(* IEC 61131-3 sources: PLC-IsaVODE/PLC-IsaVODE/samples/plc-programs (part 13) *)

(* ---- 727-SNTP_CLIENT.ST ---- *)
TYPE
  oscat_IP_FIFO128_DATA  : ARRAY [1..128] OF BYTE;
  oscat_Mailbox  : ARRAY [1..16] OF BYTE;

  oscat_IP_FIFO_DATA :
  STRUCT
    X       : oscat_IP_FIFO128_DATA; (* IP_ID FIFO Speicher          *)
    Y       : oscat_IP_FIFO128_DATA; (* IP_ID Z�hler                 *)
    ID      : BYTE;                  (* h�chste vergabene id         *)
    MAX_ID  : BYTE;                  (* maximal Anmeldungen pro ID   *)
      INIT    : BOOL;                  (* Initialisierung durchgef�hrt *)
    EMPTY   : BOOL;                  (* FIFO leer                    *)
    FULL    : BOOL;                  (* FIFO voll                    *)
    TOP     : INT;                   (* maximale anzahl in FIFO      *)
    NW      : INT;                   (* Schreibzeiger                *)
    NR      : INT;                   (* Lesezeiger                   *)
  END_STRUCT;

  oscat_IP_C:
  STRUCT
    C_MODE:			BYTE;          		(*W Mode: TCP/UCP AKTIV/PASSIV                               *)
    C_PORT:         WORD;          		(*W Portnummer                                               *)
    C_IP:           DWORD;         		(*W IP-Adresse gepackt wwxxyyzz = www.xxx.yyy.zzz            *)
    C_STATE:        BYTE;          		(*R Verbindungsstatus ON/OFF + Flanke ON/OFF                 *)
    C_ENABLE:       BOOL;          		(*W Freigabe f�r Connect                                     *)
    R_OBSERVE:      BOOL;          		(*W Empfang ueberwachen                                      *)
    TIME_RESET:     BOOL;          		(*W Alle Timer ruecksetzen                                   *)
    ERROR:          DWORD;         		(*R vvwwxxyy (vv = CON_ERROR, ww = SEN_ERROR, xx = REC_ERROR *)
    FIFO:           oscat_IP_FIFO_DATA; (*I IP FIFO Struktur                                         *)
    MAILBOX:		oscat_Mailbox;		(*I Mailbox: Datenbereich f�r Bausteindatenaustausch         *)
  END_STRUCT;
END_TYPE

TYPE

  oscat_NW_BUF_LONG  : ARRAY [0..4095] OF BYTE;

  oscat_NETWORK_BUFFER :
  STRUCT
    SIZE   : UINT;
    BUFFER : oscat_NW_BUF_LONG;
  END_STRUCT;

END_TYPE

FUNCTION _BYTE_TO_INT:INT
	VAR_INPUT
		IN :	BYTE;
	END_VAR

	_BYTE_TO_INT := USINT_TO_INT(BYTE_TO_USINT(IN));
END_FUNCTION

FUNCTION_BLOCK IP_FIFO_Block

  VAR_IN_OUT
    FIFO :	oscat_IP_FIFO_DATA;
    ID :	BYTE;
    STATE :	BYTE;
  END_VAR

  VAR
    tmp :	INT;
  END_VAR

  IF NOT FIFO.INIT THEN
    FIFO.INIT		:= TRUE;
    FIFO.NW		:= 1;
    FIFO.NR		:= 1;
    FIFO.EMPTY	:= TRUE;
    FIFO.FULL		:= FALSE;
    FIFO.TOP		:= 128;
    FIFO.MAX_ID	:= BYTE#1;
  END_IF;

  IF ID = BYTE#00 THEN
    IF FIFO.ID < INT_TO_BYTE(FIFO.TOP) THEN
      ID := USINT_TO_BYTE(BYTE_TO_USINT(FIFO.ID) + USINT#1);
      FIFO.ID := ID ;

    ELSIF STATE < BYTE#200 THEN
      STATE := BYTE#255;
    RETURN;
    END_IF;
  END_IF;

  IF STATE = BYTE#1 AND NOT FIFO.FULL THEN
    tmp := _BYTE_TO_INT(ID);
    IF FIFO.Y[tmp] < FIFO.MAX_ID THEN
      FIFO.Y[tmp] := USINT_TO_BYTE(BYTE_TO_USINT(FIFO.Y[tmp]) + USINT#1);
      tmp := FIFO.NW;
      FIFO.X[tmp] := ID;
      IF FIFO.NW = FIFO.TOP THEN FIFO.NW := 1; ELSE FIFO.NW := FIFO.NW + 1; END_IF;
      FIFO.FULL := FIFO.NW = FIFO.NR;
    FIFO.EMPTY := FALSE;
      STATE := BYTE#2;
    END_IF;
  END_IF;

  IF STATE = BYTE#2 AND NOT FIFO.EMPTY THEN
    tmp := FIFO.NR;
    IF ID = FIFO.X[tmp] THEN
      STATE := BYTE#3;
    END_IF;
  END_IF;

  IF STATE = BYTE#4 AND NOT FIFO.EMPTY THEN

    tmp := FIFO.NR;
    IF ID = FIFO.X[tmp] THEN
      tmp := _BYTE_TO_INT(ID);
      FIFO.Y[tmp] := USINT_TO_BYTE(BYTE_TO_USINT(FIFO.Y[tmp]) - USINT#1);

      IF FIFO.NR = FIFO.TOP THEN FIFO.NR := 1; ELSE FIFO.NR := FIFO.NR + 1; END_IF;
      FIFO.EMPTY := FIFO.NR = FIFO.NW;
    FIFO.FULL := FALSE;
    END_IF;
    STATE := BYTE#5;
  END_IF;

END_FUNCTION_BLOCK

FUNCTION_BLOCK T_PLC_MS_block

	VAR_OUTPUT
		T_PLC_MS :	UDINT;
	END_VAR

	VAR_EXTERNAL
		PLC_TICKS_PER_SEC :	INT;
		PLC_SYS_TICK_CNT :	DINT;
	END_VAR

	VAR
		debug :	BOOL;(*Debug-Mode ON / OFF*)
		N :	INT;(*Debug-Faktor*)
		Offset :	UDINT;(*Debug-Offset*)
		temp :	DWORD := DWORD#1;(*Debug-Offset*)
		mode :	BOOL;(*modus*)
		faktor :	UDINT;(*Systemtakt-Faktor*)
		init :	BOOL;
		v_plc_ticks_per_sec :	UDINT;
		base :	UDINT := UDINT#1000;
	END_VAR

	IF init = FALSE THEN
		v_plc_ticks_per_sec := INT_TO_UDINT(PLC_TICKS_PER_SEC);
		IF v_plc_ticks_per_sec = UDINT#1024 THEN
			faktor := UDINT#1;
			mode := FALSE;
		ELSIF v_plc_ticks_per_sec > UDINT#0 THEN
			IF v_plc_ticks_per_sec <= base THEN
				faktor := base / v_plc_ticks_per_sec;
				mode := FALSE;
			ELSE
				faktor := v_plc_ticks_per_sec / base;
				mode := TRUE;
			END_IF;
		ELSE
			faktor := UDINT#1;
		END_IF;
		init := TRUE;
	END_IF;

	IF mode THEN
		T_PLC_MS := DINT_TO_UDINT(PLC_SYS_TICK_CNT) / faktor;
	ELSE
		T_PLC_MS := DINT_TO_UDINT(PLC_SYS_TICK_CNT) * faktor;
	END_IF;

	IF debug THEN
		T_PLC_MS := (DWORD_TO_UDINT(SHL(UDINT_TO_DWORD(T_PLC_MS),N) OR SHL(temp,N)) - UDINT#1) + Offset;
	END_IF;

END_FUNCTION_BLOCK

FUNCTION DWORD_OF_BYTE:DWORD
	VAR_INPUT
		B3 :	BYTE;
		B2 :	BYTE;
		B1 :	BYTE;
		B0 :	BYTE;
	END_VAR

	DWORD_OF_BYTE := SHL(SHL(SHL(BYTE_TO_DWORD(B3),8) OR BYTE_TO_DWORD(B2),8) OR BYTE_TO_DWORD(B1),8) OR BYTE_TO_DWORD(B0);

END_FUNCTION

FUNCTION _WORD_TO_DINT:DINT
	VAR_INPUT
		IN :	WORD;
	END_VAR
	_WORD_TO_DINT := UINT_TO_DINT(WORD_TO_UINT(IN));
END_FUNCTION

FUNCTION WORD_OF_BYTE:WORD
	VAR_INPUT
		B1 :	BYTE;
		B0 :	BYTE;
	END_VAR
	WORD_OF_BYTE := SHL(BYTE_TO_WORD(B1),8) OR BYTE_TO_WORD(B0);
END_FUNCTION

FUNCTION _INT_TO_UDINT:UDINT
	VAR_INPUT
		IN :	INT;
	END_VAR

	_INT_TO_UDINT := DINT_TO_UDINT(INT_TO_DINT(IN));
END_FUNCTION

FUNCTION_BLOCK SNTP_CLIENT_Block

  VAR_IN_OUT
    IP_C :	oscat_IP_C;
    S_BUF :	oscat_NETWORK_BUFFER;
    R_BUF :	oscat_NETWORK_BUFFER;
  END_VAR

  VAR_INPUT
    IP4 :	DWORD;
    ACTIVATE :	BOOL;
  END_VAR

  VAR_OUTPUT
    ERROR :	DWORD;
    DONE_P :	BOOL;
    UDT :	UDINT;
    XMS :	INT;
  END_VAR

  VAR
    IP_STATE :	BYTE;
    IP_ID :	BYTE;
    IP_FIFO :	IP_FIFO_Block;
    i :	INT;
    last :	UDINT;
    state :	INT;
    T_PLC_MS :	T_PLC_MS_Block;
    tx :	UDINT;
    ACTIVATE_LAST :	BOOL;
    IP4_STORED :	DWORD;
  END_VAR

  T_PLC_MS();
  tx := T_PLC_MS.T_PLC_MS;

  CASE state OF
  00:
    DONE_P := FALSE;
    IF ACTIVATE AND NOT ACTIVATE_LAST THEN
      IP4_STORED := IP4;
      state := 10;
      ERROR := DWORD#0;
      IP_STATE := BYTE#1;
    END_IF;

  10:
    IF IP_STATE = BYTE#3 THEN

      S_BUF.BUFFER[00] := BYTE#16#1B;
      FOR i := 1 TO 47 DO
        S_BUF.BUFFER[i] := BYTE#16#00;
      END_FOR;

      last := tx;
      state := 30;

      IP_C.C_PORT     := WORD#123;
      IP_C.C_IP       := IP4_STORED;
      IP_C.C_MODE     := BYTE#1;
      IP_C.C_ENABLE   := TRUE;
      IP_C.TIME_RESET := TRUE;
      IP_C.R_OBSERVE  := TRUE;
      S_BUF.SIZE      := UINT#48;
      R_BUF.SIZE      := UINT#0;
    END_IF;

  30:
    IF IP_C.ERROR <> DWORD#00 THEN
      ERROR := IP_C.ERROR;
    S_BUF.SIZE := UINT#0;
    R_BUF.SIZE := UINT#0;
      state := 0;
    ELSIF S_BUF.SIZE = UINT#0 AND R_BUF.SIZE >= UINT#48 THEN
      UDT := DWORD_TO_UDINT(DWORD_OF_BYTE(R_BUF.BUFFER[40],R_BUF.BUFFER[41],R_BUF.BUFFER[42],R_BUF.BUFFER[43]))- UDINT#2208988800;

      XMS := DWORD_TO_INT(SHR(DINT_TO_DWORD(_WORD_TO_DINT(WORD_OF_BYTE(R_BUF.BUFFER[44],R_BUF.BUFFER[45])) * DINT#1000),16));
      XMS := XMS + DWORD_TO_INT(SHR(UDINT_TO_DWORD(tx - last),1));

      UDT := UDT + _INT_TO_UDINT(XMS / 1000);
      XMS := XMS MOD 1000;

      state := 0;
      DONE_P := TRUE;

    END_IF;

    IF state = 0 THEN
      IP_C.R_OBSERVE := FALSE;
      IP_STATE := BYTE#4;
    END_IF;

  END_CASE;

  ACTIVATE_LAST := ACTIVATE;

  IP_FIFO(FIFO:=IP_C.FIFO,STATE:=IP_STATE,ID:=IP_ID);
  IP_C.FIFO:=IP_FIFO.FIFO;
  IP_STATE := IP_FIFO.STATE;
  IP_ID:=IP_FIFO.ID;

END_FUNCTION_BLOCK

PROGRAM program0
	VAR
		IP_C :	oscat_IP_C;
    S_BUF :	oscat_NETWORK_BUFFER;
    R_BUF :	oscat_NETWORK_BUFFER;
    IP4 :	DWORD;
    ACTIVATE :	BOOL;
    ERROR :	DWORD;
    DONE_P :	BOOL;
    UDT :	UDINT;
    XMS :	INT;

		func_block : SNTP_CLIENT_Block;
	END_VAR
	func_block.IP_C := IP_C;
	func_block.S_BUF := S_BUF;
	func_block.R_BUF := R_BUF;
  func_block.IP4 := IP4;
	func_block.ACTIVATE := ACTIVATE;

	func_block();
  IP_C  := func_block.IP_C;
  S_BUF  := func_block.S_BUF;
  R_BUF  := func_block.R_BUF;
  ERROR  := func_block.ERROR;
  DONE_P  := func_block.DONE_P;
  UDT  := func_block.UDT;
  XMS  := func_block.XMS;
END_PROGRAM

CONFIGURATION Config0

	VAR_GLOBAL
		PLC_TICKS_PER_SEC :	INT;
		PLC_SYS_TICK_CNT :	DINT;
	END_VAR

  	RESOURCE Res0 ON PLC
    	TASK task0(INTERVAL := T#20ms,PRIORITY := 0);
    	PROGRAM instance0 WITH task0 : program0;
  	END_RESOURCE

END_CONFIGURATION

(* ---- 728-HOLIDAY.ST ---- *)
TYPE oscat_LANGUAGE:
  STRUCT
    DEFAULT 	: INT;
	LMAX    	: INT;
  END_STRUCT;
END_TYPE

TYPE
	oscat_LOCATION_ELEMENTS	: ARRAY [1..5] OF INT;
END_TYPE

TYPE
  oscat_ELEMENT_WEEKDAYS	: ARRAY [1..7] OF STRING;
  oscat_WEEKDAYS			: ARRAY [1..3]  OF oscat_ELEMENT_WEEKDAYS := [0, 0, 0];
END_TYPE

TYPE oscat_LOCATION:
  STRUCT
    DEFAULT 	: INT;
	LMAX    	: INT;
	LANGUAGE	: oscat_LOCATION_ELEMENTS;
  END_STRUCT;
END_TYPE

TYPE oscat_HOLIDAY_DATA :
  STRUCT
	NAME : STRING;
	DAY : SINT;
	MONTH : SINT;
	USE : SINT;
	PAD_BYTE : BYTE;
  END_STRUCT;
END_TYPE

TYPE
  oscat_HOLIDAY_DATA_0_29 	: ARRAY [0..29] OF oscat_HOLIDAY_DATA;
  oscat_HOLIDAY_DATA_0_49 	: ARRAY [0..49] OF oscat_HOLIDAY_DATA;
END_TYPE

FUNCTION_BLOCK SETUP_LANGUAGE_Block

	VAR_IN_OUT
		LANGUAGE :	oscat_LANGUAGE;
	END_VAR

	VAR
		init :	BOOL;
	END_VAR

	IF init THEN RETURN; END_IF;
	init := TRUE;

	LANGUAGE.DEFAULT  := 1; (* 1=english, 2=german 3=french *)
	LANGUAGE.LMAX := 3;
END_FUNCTION_BLOCK

FUNCTION_BLOCK SETUP_LOCATION
	VAR_IN_OUT
		LOCATION :	oscat_LOCATION;
	END_VAR

	VAR
		init :	BOOL;
	END_VAR

	IF init THEN RETURN; END_IF;
	init := TRUE;

	LOCATION.DEFAULT  := 1;
	LOCATION.LMAX := 5;

	LOCATION.LANGUAGE[1] := 2;
	LOCATION.LANGUAGE[2] := 2;
	LOCATION.LANGUAGE[3] := 3;
	LOCATION.LANGUAGE[4] := 2;
	LOCATION.LANGUAGE[5] := 2;
END_FUNCTION_BLOCK

FUNCTION_BLOCK SETUP_WEEKDAYS

	VAR_IN_OUT
		WEEKDAYS :	oscat_WEEKDAYS;
	END_VAR

	VAR
		init :	BOOL;
	END_VAR

	IF init THEN RETURN; END_IF;
	init := TRUE;

	WEEKDAYS[1][01] := 'Monday';
	WEEKDAYS[1][02] := 'Tuesday';
	WEEKDAYS[1][03] := 'Wednesday';
	WEEKDAYS[1][04] := 'Thursday';
	WEEKDAYS[1][05] := 'Friday';
	WEEKDAYS[1][06] := 'Saturday';
	WEEKDAYS[1][07] := 'Sunday';

	WEEKDAYS[2][01] := 'Montag';
	WEEKDAYS[2][02] := 'Dienstag';
	WEEKDAYS[2][03] := 'Mittwoch';
	WEEKDAYS[2][04] := 'Donnerstag';
	WEEKDAYS[2][05] := 'Freitag';
	WEEKDAYS[2][06] := 'Samstag';
	WEEKDAYS[2][07] := 'Sonntag';

	WEEKDAYS[3][01] := 'Lundi';
	WEEKDAYS[3][02] := 'Mardi';
	WEEKDAYS[3][03] := 'Mercredi';
	WEEKDAYS[3][04] := 'Jeudi';
	WEEKDAYS[3][05] := 'Vendredi';
	WEEKDAYS[3][06] := 'Samedi';
	WEEKDAYS[3][07] := 'Dimanche';
END_FUNCTION_BLOCK

FUNCTION YEAR_OF_DATE:INT
	VAR_INPUT
		IDATE :	UDINT;
	END_VAR

	YEAR_OF_DATE := UDINT_TO_INT((idate+UDINT#43200) / UDINT#31557600 + UDINT#1970);
END_FUNCTION

FUNCTION _INT_TO_UDINT:UDINT
	VAR_INPUT
		IN :	INT;
	END_VAR

	_INT_TO_UDINT := DINT_TO_UDINT(INT_TO_DINT(IN));
END_FUNCTION

FUNCTION SET_DATE:UDINT

	VAR_INPUT
		YEAR :	INT;
		MONTH :	INT;
		DAY :	INT;
	END_VAR

	VAR
		count :	INT;
	END_VAR

	IF month > 2 THEN
		count := (month - 1) * 30;
		IF month > 7 THEN
			count := count + DWORD_TO_INT(SHR(DINT_TO_DWORD(INT_TO_DINT(month) - INT_TO_DINT(3)),1));
		ELSE
			count := count + DWORD_TO_INT(SHR(DINT_TO_DWORD(INT_TO_DINT(month) - INT_TO_DINT(4)),1));
		END_IF;
		IF SHL(INT_TO_WORD(year),14) = WORD#0 THEN
			count := count + 1;
		END_IF;
	ELSE
		count := (month - 1) * 31;
	END_IF;
	SET_DATE := (_INT_TO_UDINT(count + day - 1) + DWORD_TO_UDINT(SHR(UDINT_TO_DWORD(_INT_TO_UDINT(year) * UDINT#1461 - UDINT#2878169), 2))) * UDINT#86400;
END_FUNCTION

FUNCTION DAY_OF_WEEK:INT
	VAR_INPUT
		IDATE :	UDINT;
	END_VAR

	DAY_OF_WEEK := UDINT_TO_INT((idate / UDINT#86400 + UDINT#3) MOD UDINT#7) + INT#01;
END_FUNCTION

FUNCTION EASTER:UDINT
	VAR_INPUT
		YEAR :	INT;
	END_VAR

	VAR
		b :	INT;
		c :	INT;
		oday :	INT;
	END_VAR

	b := (204 - 11 * (year MOD 19)) MOD 30;
	IF b > 27 THEN b := b - 1; END_IF;
	c := (year + WORD_TO_INT(SHR(INT_TO_WORD(year),2)) + b - 13) MOD 7;
	oday := 28 + b - c;
	IF oday > 33 THEN
		easter := set_Date(year, 4, oday - 31);
	ELSE
		easter := set_Date(year, 3, oday);
	END_IF;
END_FUNCTION

FUNCTION LEAP_OF_DATE:BOOL

	VAR_INPUT
		IDATE :	UDINT;
	END_VAR

	LEAP_OF_DATE := SHL(UDINT_TO_DWORD((idate + UDINT#43200) / UDINT#31557600), 30) = DWORD#16#80000000;
END_FUNCTION

FUNCTION DAY_OF_YEAR:INT
	VAR_INPUT
		IDATE :	UDINT;
	END_VAR

	DAY_OF_YEAR := UDINT_TO_INT(((idate) / UDINT#86400) MOD UDINT#1461);
	IF DAY_OF_YEAR > 729 THEN
		IF DAY_OF_YEAR > 1095 THEN DAY_OF_YEAR := DAY_OF_YEAR - 1095; ELSE DAY_OF_YEAR := DAY_OF_YEAR - 729; END_IF;
	ELSIF DAY_OF_YEAR > 364 THEN
		DAY_OF_YEAR := DAY_OF_YEAR - 364;
	ELSE
		DAY_OF_YEAR := DAY_OF_YEAR + 1;
	END_IF;
END_FUNCTION

FUNCTION MONTH_OF_DATE:INT

	VAR_INPUT
		IDATE :	UDINT;
	END_VAR

	MONTH_OF_DATE := DAY_OF_YEAR(idate);
	IF MONTH_OF_DATE < 32 THEN
		MONTH_OF_DATE := 1;
	ELSIF LEAP_OF_DATE((IDATE)) THEN
		MONTH_OF_DATE := (MONTH_OF_DATE * 53 + 1668) / 1623;
	ELSE
		MONTH_OF_DATE := (MONTH_OF_DATE * 53 + 1700) / 1620;
	END_IF;
END_FUNCTION

FUNCTION DAY_OF_MONTH:INT
	VAR_INPUT
		IDATE :	UDINT;
	END_VAR

	day_of_month := day_of_year(idate);

	IF leap_of_Date((idate)) THEN
		CASE day_of_month OF
			32..60	:	day_of_month := day_of_month - 31;
			61..91	:	day_of_month := day_of_month - 60;
			92..121 :	day_of_month := day_of_month - 91;
			122..152:	day_of_month := day_of_month - 121;
			153..182:	day_of_month := day_of_month - 152;
			183..213:	day_of_month := day_of_month - 182;
			214..244:	day_of_month := day_of_month - 213;
			245..274:	day_of_month := day_of_month - 244;
			275..305:	day_of_month := day_of_month - 274;
			306..335:	day_of_month := day_of_month - 305;
			336..366:	day_of_month := day_of_month - 335;
		END_CASE;
	ELSE
		CASE day_of_month OF
			32..59	:	day_of_month := day_of_month - 31;
			60..90	:	day_of_month := day_of_month - 59;
			91..120 :	day_of_month := day_of_month - 90;
			121..151:	day_of_month := day_of_month - 120;
			152..181:	day_of_month := day_of_month - 151;
			182..212:	day_of_month := day_of_month - 181;
			213..243:	day_of_month := day_of_month - 212;
			244..273:	day_of_month := day_of_month - 243;
			274..304:	day_of_month := day_of_month - 273;
			305..334:	day_of_month := day_of_month - 304;
			335..365:	day_of_month := day_of_month - 334;
		END_CASE;
	END_IF;
END_FUNCTION

FUNCTION DATE_ADD:UDINT
	VAR_INPUT
		IDATE :	UDINT;
		D :	INT;
		W :	INT;
		M :	INT;
		Y :	INT;
	END_VAR

	VAR
		mo :	INT;
		yr :	INT;
		dm :	INT;
	END_VAR

	DATE_ADD := IDATE + INT_TO_UDINT(D + W * 7) * UDINT#86400;
	yr := Y + YEAR_OF_DATE(DATE_ADD);
	mo := M + MONTH_OF_DATE(DATE_ADD);
	dm := DAY_OF_MONTH(DATE_ADD);
	WHILE mo > 12 DO
		mo := mo - 12;
		yr := yr + 1;
	END_WHILE;
	WHILE mo < 1 DO
		mo := mo + 12;
		yr := yr - 1;
	END_WHILE;
	DATE_ADD := SET_DATE(yr, mo, dm);
END_FUNCTION

FUNCTION_BLOCK HOLIDAY_Block
	VAR_INPUT
		DATE_IN :	UDINT;
		LANGU :	INT;
		FRIDAY :	BOOL;
		SATURDAY :	BOOL;
		SUNDAY :	BOOL;
	END_VAR

	VAR_IN_OUT
		HOLIDAYS :	oscat_HOLIDAY_DATA_0_29;
	END_VAR

	VAR_OUTPUT
		Y :	BOOL;
		NAME :	STRING;
	END_VAR

	VAR
		size :	INT := INT#29;
		last_active :	UDINT;
		ostern :	UDINT;
		i :	INT;
		jahr :	INT;
		x_date :	UDINT;
		lx :	INT;
		wdx :	INT;
		SETUP_LOCATIONS :	SETUP_LOCATION;
		SETUP_WEEKDAYSS :	SETUP_WEEKDAYS;
		SETUP_LANGUAGES :	SETUP_LANGUAGE_Block;
		LOCATION :	oscat_LOCATION;
		WEEKDAYS :	oscat_WEEKDAYS;
		LANGUAGE :	oscat_LANGUAGE;
		wd :	INT;
	END_VAR

	IF last_active = date_in THEN RETURN; END_IF;
	last_active := DATE_IN;

	SETUP_LOCATIONS(LOCATION:=LOCATION);
	LOCATION:=SETUP_LOCATIONS.LOCATION;

	SETUP_WEEKDAYSS(WEEKDAYS:=WEEKDAYS);
	WEEKDAYS:=SETUP_WEEKDAYSS.WEEKDAYS;

	SETUP_LANGUAGES(LANGUAGE:=LANGUAGE);
	LANGUAGE:=SETUP_LANGUAGES.LANGUAGE;

	IF LANGU = 0 THEN
		lx := language.DEFAULT;
	ELSE
		lx := MIN(language.LMAX, LANGU);
	END_IF;

	jahr := YEAR_OF_DATE(date_in);
	ostern := EASTER(jahr);
	wdx := DAY_OF_WEEK(DATE_IN);
	Y := FALSE;

	FOR i := 0 TO size DO
		x_date := SET_DATE(jahr, SINT_TO_INT(HOLIDAYS[i].MONTH) , SINT_TO_INT(HOLIDAYS[i].DAY));
		IF HOLIDAYS[i].USE = SINT#1 AND HOLIDAYS[i].MONTH > SINT#0 THEN
			(* check for fixed date holiday *)
			IF x_date = date_in THEN
				Y := TRUE;
				NAME := HOLIDAYS[i].NAME;
				RETURN;
			END_IF;
		ELSIF HOLIDAYS[i].USE = SINT#1 AND HOLIDAYS[i].MONTH = SINT#0 THEN
			(* check for holiday in reference to easter *)
			IF DATE_ADD(ostern, SINT_TO_INT(HOLIDAYS[i].DAY),0,0,0) = date_in THEN
				Y := TRUE;
				NAME := HOLIDAYS[i].NAME;
				RETURN;
			END_IF;
		ELSIF HOLIDAYS[i].USE < SINT#0 THEN
			(* check for holiday on a weekday before date *)
			IF DAY_OF_WEEK(date_in) = SINT_TO_INT(ABS(HOLIDAYS[i].USE)) AND date_in < x_date AND date_in >= DATE_ADD(x_date,-7,0,0,0) THEN
				Y := TRUE;
				NAME := HOLIDAYS[i].NAME;
				RETURN;
			END_IF;
		END_IF;
	END_FOR;

	IF NOT Y AND (wdx = 5 AND FRIDAY OR wdx = 6 AND SATURDAY OR wdx = 7 AND SUNDAY) THEN
		Y := TRUE;
		wd := LOCATION.LANGUAGE[lx];
		NAME := WEEKDAYS[wd][wdx];
	ELSE
		NAME := '';
	END_IF;
END_FUNCTION_BLOCK

PROGRAM program0
  VAR
	DATE_IN  :	UDINT;
	LANGU    :	INT;
	FRIDAY   :	BOOL;
	SATURDAY :	BOOL;
	SUNDAY   :	BOOL;

	Y :	BOOL;
	NAME :	STRING;

	HOLIDAYS :	oscat_HOLIDAY_DATA_0_29;

	func_block : HOLIDAY_Block;
  END_VAR
	func_block.DATE_IN :=DATE_IN ;
	func_block.LANGU   :=LANGU   ;
	func_block.FRIDAY  :=FRIDAY  ;
	func_block.SATURDAY:=SATURDAY;
	func_block.SUNDAY  :=SUNDAY  ;
	func_block.HOLIDAYS  :=HOLIDAYS ;

	func_block();
	Y := func_block.Y;
	NAME := func_block.NAME;
	HOLIDAYS := func_block.HOLIDAYS;

END_PROGRAM

CONFIGURATION Config0
  RESOURCE Res0 ON PLC
    TASK task0(INTERVAL := T#20ms,PRIORITY := 0);
    PROGRAM instance0 WITH task0 : program0;
  END_RESOURCE
END_CONFIGURATION

(* ---- 732-LEGIONELLA.ST ---- *)
FUNCTION TIMECHECK:BOOL

	VAR_INPUT
		TD :	UDINT;
		START :	UDINT;
		STOP :	UDINT;
	END_VAR

	IF stop < start THEN
		TIMECHECK := start <= TD OR  TD < stop;
	ELSE
		TIMECHECK := start <= TD AND TD < stop;
	END_IF;

END_FUNCTION

FUNCTION TIME_TO_TOD:UDINT

	VAR_INPUT
		IN :	TIME;
	END_VAR

	TIME_TO_TOD := DWORD_TO_UDINT(TIME_TO_DWORD(IN));
END_FUNCTION

FUNCTION TOD_TO_TIME:TIME
	VAR_INPUT
		IN :	UDINT;
	END_VAR

	TOD_TO_TIME := DWORD_TO_TIME(UDINT_TO_DWORD(IN));
END_FUNCTION

FUNCTION DAY_OF_WEEK:INT
  VAR_INPUT
    IDATE :	UDINT;
  END_VAR

  DAY_OF_WEEK := UDINT_TO_INT((idate / UDINT#86400 + UDINT#3) MOD UDINT#7) + INT#01;
END_FUNCTION

FUNCTION _DT_TO_DATE_B:UDINT

	VAR_INPUT
		_INN :	UDINT;
	END_VAR

	_DT_TO_DATE_B := (_INN / UDINT#86400) * UDINT#86400;
END_FUNCTION

FUNCTION DT_TO_TOD2:UDINT
	VAR_INPUT
		IN :	UDINT;
	END_VAR

	DT_TO_TOD2 := (IN MOD UDINT#86400) * UDINT#1000;
END_FUNCTION

FUNCTION TIME_TO_TOD2:UDINT

	VAR_INPUT
		IN :	TIME;
	END_VAR

	TIME_TO_TOD2 := DWORD_TO_UDINT(TIME_TO_DWORD(IN));
END_FUNCTION

FUNCTION_BLOCK TIMER_1_Block

	VAR_INPUT
		E :	BOOL := TRUE;
		DTI :	UDINT;
		START :	UDINT;
		DURATION :	TIME;
		DAY :	BYTE := BYTE#2#0111_1111;
	END_VAR

	VAR_OUTPUT
		Q :	BOOL;
		STOP :	TIME;
	END_VAR

	IF E THEN
		stop := TOD_TO_TIME(START) + DURATION;
		IF stop > T#24h THEN stop := stop - T#24h; END_IF;
		Q := TIMECHECK(DT_TO_TOD2(DTI), START, TIME_TO_TOD2(stop)) AND (SHR(BYTE#128, DAY_OF_WEEK(_DT_TO_DATE_B(DTI))) AND DAY) > BYTE#0;
	ELSE
		Q := FALSE;
	END_IF;

END_FUNCTION_BLOCK

FUNCTION UDINT_TO_TIME2:TIME

	VAR_INPUT
		IN :	UDINT;
	END_VAR

	UDINT_TO_TIME2 := DINT_TO_TIME(UDINT_TO_DINT(IN));

END_FUNCTION

FUNCTION_BLOCK T_PLC_MS_block
	VAR_OUTPUT
		T_PLC_MS :	UDINT;
	END_VAR

	VAR_EXTERNAL
		PLC_TICKS_PER_SEC :	INT;
		PLC_SYS_TICK_CNT :	DINT;
	END_VAR

	VAR
		debug :	BOOL;
		N :	INT;
		Offset :	UDINT;
		temp :	DWORD := DWORD#1;
		mode :	BOOL;
		faktor :	UDINT;
		init :	BOOL;
		v_plc_ticks_per_sec :	UDINT;
		base :	UDINT := UDINT#1000;
	END_VAR

	IF init = FALSE THEN
		v_plc_ticks_per_sec := INT_TO_UDINT(PLC_TICKS_PER_SEC);
		IF v_plc_ticks_per_sec = UDINT#1024 THEN
			faktor := UDINT#1;
			mode := FALSE;
		ELSIF v_plc_ticks_per_sec > UDINT#0 THEN
			IF v_plc_ticks_per_sec <= base THEN
				faktor := base / v_plc_ticks_per_sec;
				mode := FALSE;
			ELSE
				faktor := v_plc_ticks_per_sec / base;
				mode := TRUE;
			END_IF;
		ELSE
			faktor := UDINT#1;
		END_IF;
		init := TRUE;
	END_IF;

	IF mode THEN
		T_PLC_MS := DINT_TO_UDINT(PLC_SYS_TICK_CNT) / faktor;
	ELSE
		T_PLC_MS := DINT_TO_UDINT(PLC_SYS_TICK_CNT) * faktor;
	END_IF;

	IF debug THEN
		T_PLC_MS := (DWORD_TO_UDINT(SHL(UDINT_TO_DWORD(T_PLC_MS),N) OR SHL(temp,N)) - UDINT#1) + Offset;
	END_IF;

END_FUNCTION_BLOCK

FUNCTION_BLOCK SEQUENCE_8_Block

	VAR_INPUT
		IN0 :	BOOL := TRUE;
		IN1 :	BOOL := TRUE;
		IN2 :	BOOL := TRUE;
		IN3 :	BOOL := TRUE;
		IN4 :	BOOL := TRUE;
		IN5 :	BOOL := TRUE;
		IN6 :	BOOL := TRUE;
		IN7 :	BOOL := TRUE;
		START :	BOOL;
		RST :	BOOL;
		WAIT0 :	TIME;
		DELAY0 :	TIME;
		WAIT1 :	TIME;
		DELAY1 :	TIME;
		WAIT2 :	TIME;
		DELAY2 :	TIME;
		WAIT3 :	TIME;
		DELAY3 :	TIME;
		WAIT4 :	TIME;
		DELAY4 :	TIME;
		WAIT5 :	TIME;
		DELAY5 :	TIME;
		WAIT6 :	TIME;
		DELAY6 :	TIME;
		WAIT7 :	TIME;
		DELAY7 :	TIME;
		STOP_ON_ERROR :	BOOL;
	END_VAR

	VAR_OUTPUT
		Q0 :	BOOL;
		Q1 :	BOOL;
		Q2 :	BOOL;
		Q3 :	BOOL;
		Q4 :	BOOL;
		Q5 :	BOOL;
		Q6 :	BOOL;
		Q7 :	BOOL;
		QX :	BOOL;
		RUN :	BOOL;
		_STEP :	INT := -1;
		STATUS :	BYTE;
	END_VAR

	VAR
		last :	TIME;
		edge :	BOOL;
		tx :	TIME;
		init :	BOOL;
		T_PLC_MS :	T_PLC_MS_Block;
	END_VAR

	T_PLC_MS();
	tx:= UDINT_TO_TIME(T_PLC_MS.T_PLC_MS);

	IF NOT init THEN
		last := tx;
		init := TRUE;
		status := BYTE#110;
	END_IF;

	IF rst THEN
		_step := -1;
		Q0 := FALSE;
		Q1 := FALSE;
		Q2 := FALSE;
		Q3 := FALSE;
		Q4 := FALSE;
		Q5 := FALSE;
		Q6 := FALSE;
		Q7 := FALSE;
		status := BYTE#110;
		run := FALSE;

	ELSIF start AND NOT edge THEN
		_step := 0;
		last := tx;
		status := BYTE#111;
		Q0 := FALSE;
		Q1 := FALSE;
		Q2 := FALSE;
		Q3 := FALSE;
		Q4 := FALSE;
		Q5 := FALSE;
		Q6 := FALSE;
		Q7 := FALSE;
		run := TRUE;
	END_IF;
	edge := start;

	IF status > BYTE#0 AND status < BYTE#100 AND stop_on_error THEN RETURN; END_IF;

	IF run AND _step = 0 THEN
		IF NOT q0 AND in0 AND tx - last <= wait0 THEN
			Q0 := TRUE;
			last := tx;
		ELSIF NOT q0 AND tx - last > wait0 THEN
			status := BYTE#1;
			run := FALSE;
		ELSIF q0 AND tx - last >= delay0 THEN
			_step := 1;
			last := tx;
		END_IF;
	END_IF;
	IF run AND _step = 1 THEN
		IF NOT q1 AND in1 AND tx - last <= wait1 THEN
			Q0 := FALSE;
			Q1 := TRUE;
			last := tx;
		ELSIF NOT q1 AND Tx - last > wait1 THEN
			status := BYTE#2;
			q0 := FALSE;
			run := FALSE;
		ELSIF q1 AND tx - last >= delay1 THEN
			_step := 2;
			last := tx;
		END_IF;
	END_IF;
	IF run AND _step = 2 THEN
		IF NOT q2 AND in2 AND tx - last <= wait2 THEN
			Q1 := FALSE;
			Q2 := TRUE;
			last := tx;
		ELSIF NOT q2 AND Tx - last > wait2 THEN
			status := BYTE#3;
			q1 := FALSE;
			run := FALSE;
		ELSIF q2 AND tx - last >= delay2 THEN
			_step := 3;
			last := tx;
		END_IF;
	END_IF;
	IF run AND _step = 3 THEN
		IF NOT q3 AND in3 AND tx - last <= wait3 THEN
			Q2 := FALSE;
			Q3 := TRUE;
			last := tx;
		ELSIF NOT q3 AND Tx - last > wait3 THEN
			status := BYTE#4;
			q2 := FALSE;
			run := FALSE;
		ELSIF q3 AND tx - last >= delay3 THEN
			_step := 4;
			last := tx;
		END_IF;
	END_IF;
	IF run AND _step = 4 THEN
		IF NOT q4 AND in4 AND tx - last <= wait4 THEN
			Q3 := FALSE;
			Q4 := TRUE;
			last := tx;
		ELSIF NOT q4 AND Tx - last > wait4 THEN
			status := BYTE#5;
			q3 := FALSE;
			run := FALSE;
		ELSIF q4 AND tx - last >= delay4 THEN
			_step := 5;
			last := tx;
		END_IF;
	END_IF;
	IF run AND _step = 5 THEN
		IF NOT q5 AND in5 AND tx - last <= wait5 THEN
			Q4 := FALSE;
			Q5 := TRUE;
			last := tx;
		ELSIF NOT q5 AND Tx - last > wait5 THEN
			status := BYTE#6;
			q4 := FALSE;
			run := FALSE;
		ELSIF q5 AND tx - last >= delay5 THEN
			_step := 6;
			last := tx;
		END_IF;
	END_IF;
	IF run AND _step = 6 THEN
		IF NOT q6 AND in6 AND tx - last <= wait6 THEN
			Q5 := FALSE;
			Q6 := TRUE;
			last := tx;
		ELSIF NOT q6 AND Tx - last > wait6 THEN
			status := BYTE#7;
			q5 := FALSE;
			run := FALSE;
		ELSIF q6 AND tx - last >= delay6 THEN
			_step := 7;
			last := tx;
		END_IF;
	END_IF;
	IF run AND _step = 7 THEN
		IF NOT q7 AND in7 AND tx - last <= wait7 THEN
			Q6 := FALSE;
			Q7 := TRUE;
			last := tx;
		ELSIF NOT q7 AND Tx - last > wait7 THEN
			status := BYTE#8;
			q6 := FALSE;
			run := FALSE;
		ELSIF q7 AND tx - last >= delay7 THEN
			_step := -1;
			Q7 := FALSE;
			Run := FALSE;
			status := BYTE#110;
		END_IF;
	END_IF;
	QX := q0 OR q1 OR q2 OR q3 OR q4 OR q5 OR q6 OR q7;

END_FUNCTION_BLOCK

FUNCTION_BLOCK HYST_1_Block

	VAR_INPUT
		IN :	REAL;
		HIGH :	REAL;
		LOW :	REAL;
	END_VAR

	VAR_OUTPUT
		Q :	BOOL;
		WIN :	BOOL;
	END_VAR

	IF in < low THEN
		Q := FALSE;
		win := FALSE;
	ELSIF in > high THEN
		Q := TRUE;
		win := FALSE;
	ELSE
		win := TRUE;
	END_IF;

END_FUNCTION_BLOCK

FUNCTION_BLOCK LEGIONELLA_Block

	VAR_INPUT
		MANUAL :	BOOL;
		TEMP_BOILER :	REAL;
		TEMP_RETURN :	REAL := 100.0;
		DT_IN :	UDINT;
		RST :	BOOL;
		T_START :	UDINT := UDINT#10800000;(*tod#03:00:00*)
		DAY :	INT := 7;
		TEMP_SET :	REAL := 70.0;
		TEMP_OFFSET :	REAL := 10.0;
		TEMP_HYS :	REAL := 5.0;
		T_MAX_HEAT :	TIME := t#10m;
		T_MAX_RET :	TIME := t#10m;
		TP_0 :	TIME := t#5m;
		TP_1 :	TIME := t#5m;
		TP_2 :	TIME := t#5m;
		TP_3 :	TIME := t#5m;
		TP_4 :	TIME := t#5m;
		TP_5 :	TIME := t#5m;
		TP_6 :	TIME := t#5m;
		TP_7 :	TIME := t#5m;
	END_VAR

	VAR_OUTPUT
		HEAT :	BOOL;
		PUMP :	BOOL;
		VALVE0 :	BOOL;
		VALVE1 :	BOOL;
		VALVE2 :	BOOL;
		VALVE3 :	BOOL;
		VALVE4 :	BOOL;
		VALVE5 :	BOOL;
		VALVE6 :	BOOL;
		VALVE7 :	BOOL;
		RUN :	BOOL;
		_STATUS :	BYTE;
	END_VAR

	VAR
		X1 :	TIMER_1_Block;
		x2 :	SEQUENCE_8_Block;
		x3 :	HYST_1_Block;
		init :	BOOL;
	END_VAR

	IF NOT init THEN
		init := TRUE;
		X1.day := SHR(BYTE#128,day);
		X1.start := T_start;
		X3.low := Temp_offset + temp_set;
		X3.high := Temp_hys + X3.low;
		X2.wait0 := T_max_heat;
		X2.delay0 := TP_0;
		X2.delay1 := TP_1;
		X2.delay2 := TP_2;
		X2.delay3 := TP_3;
		X2.delay4 := TP_4;
		X2.delay5 := TP_5;
		X2.delay6 := TP_6;
		X2.delay7 := TP_7;
		X2.wait1 := T_max_ret;
		X2.wait2 := T_max_ret;
		X2.wait3 := T_max_ret;
		X2.wait4 := T_max_ret;
		X2.wait5 := T_max_ret;
		X2.wait6 := T_max_ret;
		X2.wait7 := T_max_ret;
		X2();
	END_IF;

	X1(DTi := DT_in);
	IF X1.Q OR MANUAL OR x2.run THEN
		X3(in := temp_boiler);
		X2.in0 := X3.Q OR x3.win;
		X2.in1 := temp_return >= temp_set;
		X2.in2 := x2.in1;
		X2.in3 := x2.in1;
		X2.in4 := x2.in1;
		X2.in5 := x2.in1;
		X2.in6 := x2.in1;
		X2.in7 := x2.in1;
		X2.rst := rst;
		X2(start := X1.Q OR MANUAL);
		run := x2.run;
		pump := x2.QX;
		Heat := NOT X3.Q AND x2.run;
		valve0 := X2.Q0;
		valve1 := X2.Q1;
		valve2 := X2.Q2;
		valve3 := X2.Q3;
		valve4 := X2.Q4;
		valve5 := X2.Q5;
		valve6 := X2.Q6;
		valve7 := X2.Q7;
		pump := X2.QX;
		_STATUS := X2.status;
	ELSE
		X2(start := FALSE);
		_STATUS := x2.status;
	END_IF;

END_FUNCTION_BLOCK

PROGRAM program0
	VAR
		MANUAL :	BOOL;
		TEMP_BOILER :	REAL;
		TEMP_RETURN :	REAL := 100.0;
		DT_IN :	UDINT;
		RST :	BOOL;
		T_START :	UDINT := UDINT#10800000;(*tod#03:00:00*)
		DAY :	INT := 7;
		TEMP_SET :	REAL := 70.0;
		TEMP_OFFSET :	REAL := 10.0;
		TEMP_HYS :	REAL := 5.0;
		T_MAX_HEAT :	TIME := t#10m;
		T_MAX_RET :	TIME := t#10m;
		TP_0 :	TIME := t#5m;
		TP_1 :	TIME := t#5m;
		TP_2 :	TIME := t#5m;
		TP_3 :	TIME := t#5m;
		TP_4 :	TIME := t#5m;
		TP_5 :	TIME := t#5m;
		TP_6 :	TIME := t#5m;
		TP_7 :	TIME := t#5m;
		HEAT :	BOOL;
		PUMP :	BOOL;
		VALVE0 :	BOOL;
		VALVE1 :	BOOL;
		VALVE2 :	BOOL;
		VALVE3 :	BOOL;
		VALVE4 :	BOOL;
		VALVE5 :	BOOL;
		VALVE6 :	BOOL;
		VALVE7 :	BOOL;
		RUN :	BOOL;
		_STATUS :	BYTE;

		func_block : LEGIONELLA_Block;
	END_VAR
	func_block.MANUAL := MANUAL;
	func_block.TEMP_BOILER := TEMP_BOILER;
	func_block.TEMP_RETURN := TEMP_RETURN ;
	func_block.DT_IN    := DT_IN    ;
	func_block.RST := RST;
	func_block.T_START := T_START;
	func_block.DAY := DAY ;
	func_block.TEMP_SET := TEMP_SET ;
	func_block.TEMP_OFFSET    := TEMP_OFFSET    ;
	func_block.TEMP_HYS    := TEMP_HYS    ;
	func_block.T_MAX_HEAT := T_MAX_HEAT;
	func_block.T_MAX_RET := T_MAX_RET;
	func_block.TP_0 := TP_0;
	func_block.TP_1 := TP_1 ;
	func_block.TP_2 := TP_2 ;
	func_block.TP_3    := TP_3    ;
	func_block.TP_4    := TP_4    ;
	func_block.TP_5 := TP_5;
	func_block.TP_6 := TP_6;
	func_block.TP_7 := TP_7;

	func_block();
	HEAT  := func_block.HEAT;
	PUMP  := func_block.PUMP;
	VALVE0  := func_block.VALVE0;
	VALVE1  := func_block.VALVE1;
	VALVE2  := func_block.VALVE2;
	VALVE3  := func_block.HEAT;
	VALVE4  := func_block.VALVE4;
	VALVE5  := func_block.VALVE5;
	VALVE6  := func_block.VALVE6;
	VALVE7  := func_block.VALVE7;
	RUN  := func_block.RUN;
	_status  := func_block._status;
END_PROGRAM

CONFIGURATION Config0
	VAR_GLOBAL
		PLC_TICKS_PER_SEC :	INT;
		PLC_SYS_TICK_CNT :	DINT;
	END_VAR
  	RESOURCE Res0 ON PLC
    	TASK task0(INTERVAL := T#20ms,PRIORITY := 0);
    	PROGRAM instance0 WITH task0 : program0;
  	END_RESOURCE
END_CONFIGURATION

(* ---- 734-DCF77.ST ---- *)
TYPE
  oscat_dcf77_bits            : ARRAY [0..58]   OF BOOL;
END_TYPE

FUNCTION_BLOCK T_PLC_MS_block
	VAR_OUTPUT
		T_PLC_MS :	UDINT;
	END_VAR

	VAR_EXTERNAL
		PLC_TICKS_PER_SEC :	INT;
		PLC_SYS_TICK_CNT :	DINT;
	END_VAR

	VAR
		debug :	BOOL;(*Debug-Mode ON / OFF*)
		N :	INT;(*Debug-Faktor*)
		Offset :	UDINT;(*Debug-Offset*)
		temp :	DWORD := DWORD#1;(*Debug-Offset*)
		mode :	BOOL;(*modus*)
		faktor :	UDINT;(*Systemtakt-Faktor*)
		init :	BOOL;
		v_plc_ticks_per_sec :	UDINT;
		base :	UDINT := UDINT#1000;
	END_VAR

	IF init = FALSE THEN
		v_plc_ticks_per_sec := INT_TO_UDINT(PLC_TICKS_PER_SEC);
		IF v_plc_ticks_per_sec = UDINT#1024 THEN
			faktor := UDINT#1;
			mode := FALSE;
		ELSIF v_plc_ticks_per_sec > UDINT#0 THEN
			IF v_plc_ticks_per_sec <= base THEN
				faktor := base / v_plc_ticks_per_sec;
				mode := FALSE;
			ELSE
				faktor := v_plc_ticks_per_sec / base;
				mode := TRUE;
			END_IF;
		ELSE
			faktor := UDINT#1;
		END_IF;
		init := TRUE;
	END_IF;

	IF mode THEN
		T_PLC_MS := DINT_TO_UDINT(PLC_SYS_TICK_CNT) / faktor;
	ELSE
		T_PLC_MS := DINT_TO_UDINT(PLC_SYS_TICK_CNT) * faktor;
	END_IF;

	IF debug THEN
		T_PLC_MS := (DWORD_TO_UDINT(SHL(UDINT_TO_DWORD(T_PLC_MS),N) OR SHL(temp,N)) - UDINT#1) + Offset;
	END_IF;

END_FUNCTION_BLOCK

FUNCTION BIT_LOAD_W:WORD
	VAR_INPUT
		IN :	WORD;
		VAL :	BOOL;
		POS :	INT;
	END_VAR

	IF VAL THEN
		BIT_LOAD_W := in OR SHL(WORD#1,pos);
	ELSE
		BIT_LOAD_W := in AND (NOT SHL(WORD#1,pos));
	END_IF;
END_FUNCTION

FUNCTION BIT_OF_DWORD:BOOL
	VAR_INPUT
		IN :	DWORD;
		N :	INT;
	END_VAR
	BIT_OF_DWORD := (SHR(in,n) AND DWORD#1) > DWORD#0;
END_FUNCTION

FUNCTION EVEN:BOOL
	VAR_INPUT
		IN :	DINT;
	END_VAR
	even := NOT BIT_OF_DWORD(DINT_TO_DWORD(in),0);
END_FUNCTION

FUNCTION _INT_TO_UDINT:UDINT
	VAR_INPUT
		IN :	INT;
	END_VAR

	_INT_TO_UDINT := DINT_TO_UDINT(INT_TO_DINT(IN));
END_FUNCTION

FUNCTION SET_DATE:UDINT

	VAR_INPUT
		YEAR :	INT;
		MONTH :	INT;
		DAY :	INT;
	END_VAR

	VAR
		count :	INT;
	END_VAR

	IF month > 2 THEN
		count := (month - 1) * 30;
		IF month > 7 THEN
			count := count + DWORD_TO_INT(SHR(DINT_TO_DWORD(INT_TO_DINT(month) - INT_TO_DINT(3)),1));
		ELSE
			count := count + DWORD_TO_INT(SHR(DINT_TO_DWORD(INT_TO_DINT(month) - INT_TO_DINT(4)),1));
		END_IF;
		IF SHL(INT_TO_WORD(year),14) = WORD#0 THEN
			count := count + 1;
		END_IF;
	ELSE
		count := (month - 1) * 31;
	END_IF;
	SET_DATE := (_INT_TO_UDINT(count + day - 1) + DWORD_TO_UDINT(SHR(UDINT_TO_DWORD(_INT_TO_UDINT(year) * UDINT#1461 - UDINT#2878169), 2))) * UDINT#86400;

END_FUNCTION

FUNCTION DST:BOOL
	VAR_INPUT
		UTC :	UDINT;
	END_VAR

	VAR
		yr :	INT;
		yr4 :	UDINT;
		ltc :	UDINT;
		idate :	UDINT;
	END_VAR

	yr := YEAR_OF_DATE(DT_TO_DATE2(UTC));
	ltc := UTC;
	idate := SET_DT(yr, 3, 31, 1, 0, 0);
	yr4 := DWORD_TO_UDINT(SHR(INT_TO_DWORD(5 * yr), 2)) + UDINT#1;
	DST := (idate - ((yr4 + UDINT#3) MOD UDINT#7) * UDINT#86400 <= ltc) AND (idate + (UDINT#214 - (yr4) MOD UDINT#7) * UDINT#86400 > ltc);

END_FUNCTION

FUNCTION YEAR_OF_DATE:INT
	VAR_INPUT
		IDATE :	UDINT;
	END_VAR

	YEAR_OF_DATE := UDINT_TO_INT((idate+UDINT#43200) / UDINT#31557600 + UDINT#1970);
END_FUNCTION

FUNCTION DAY_OF_WEEK:INT

	VAR_INPUT
		IDATE :	UDINT;
	END_VAR

	DAY_OF_WEEK := UDINT_TO_INT((idate / UDINT#86400 + UDINT#3) MOD UDINT#7) + INT#01;
END_FUNCTION

FUNCTION SET_DT:UDINT
	VAR_INPUT
		YEAR :	INT;
		MONTH :	INT;
		DAY :	INT;
		HOUR :	INT;
		MINUTE :	INT;
		SECOND :	INT;
	END_VAR

	SET_DT := SET_DATE(YEAR, MONTH, DAY) + _INT_TO_UDINT(SECOND) + _INT_TO_UDINT(MINUTE) * UDINT#60 + _INT_TO_UDINT(HOUR) * UDINT#3600;
END_FUNCTION

FUNCTION DT_TO_DATE2:UDINT

	VAR_INPUT
		IN :	UDINT;
	END_VAR

	DT_TO_DATE2 := (IN / UDINT#86400) * UDINT#86400;

END_FUNCTION

FUNCTION_BLOCK DCF77
	VAR_INPUT
		REC :	BOOL;
		SET :	BOOL;
		SDT :	UDINT;
		DSI :	BOOL;
		SYNC_TIMEOUT :	TIME := t#2m;
		TIME_OFFSET :	INT := 1;
		DST_EN :	BOOL := TRUE;
	END_VAR

	VAR_OUTPUT
		TPp :	BOOL;
		DS :	BOOL;
		WDAY :	INT;
		ERROR :	BOOL;
		RTC2 :	UDINT;
		RTC21 :	UDINT;
		MSEC :	INT;
		SYNC :	BOOL;
	END_VAR

	VAR
		MEZ :	UDINT;
		UTC :	UDINT;
		state :	INT;
		edge :	BOOL;
		tx :	TIME;
		ty :	TIME;
		last :	TIME;
		bits :	oscat_dcf77_bits;
		cnt :	INT;
		i :	INT;
		old_time :	UDINT;
		minute :	INT;
		hour :	INT;
		day :	INT;
		month :	INT;
		year :	INT;
		last_sync :	TIME;
		t1 :	TIME;
		tz :	TIME;
		init :	BOOL;
		word_temp :	WORD;
		bool_temp :	BOOL;
		T_PLC_MS :	T_PLC_MS_block;
	END_VAR

	TPp := FALSE;

	T_PLC_MS();
	t1:= UDINT_TO_TIME(T_PLC_MS.T_PLC_MS);
	tx := t1 - last;

	IF rec XOR edge THEN
		edge := rec;
		IF NOT rec AND tx > t#1700ms AND tx < t#2000ms THEN
			(* start condition reached *)
			state := 0;
			tpp := NOT error;
		ELSIF NOT rec AND tx > t#700ms AND tx < t#1000ms THEN
			(* second switch detected *)
			IF state < 58 THEN state := state +1; ELSE state := 0; END_IF;
		ELSIF rec AND tx  < t#120ms THEN
			(* bit 0 detected  *)
			bits[state] := FALSE;
		ELSIF rec AND tx > t#120ms AND tx < t#250ms THEN
			(* bit 1 detected *)
			bits[state] := TRUE;
		ELSE
			(* error condition received signal is not valid *)
			error := TRUE;
			state := 0;
		END_IF;
		last := last + tx;
		IF rec AND state = 58 THEN
			error := FALSE;

			IF bits[0] OR NOT (bits[17] XOR bits[18]) OR NOT bits[20] THEN error := TRUE; END_IF;
			word_temp := WORD#0;

			bool_temp:=bits[21];
			word_temp:=BIT_LOAD_W(word_temp,bool_temp,0);
			bool_temp:=bits[22];
			word_temp:=BIT_LOAD_W(word_temp,bool_temp,1);
			bool_temp:=bits[23];
			word_temp:=BIT_LOAD_W(word_temp,bool_temp,2);
			bool_temp:=bits[24];
			word_temp:=BIT_LOAD_W(word_temp,bool_temp,3);

			minute := WORD_TO_INT(word_temp);
			IF bits[25] THEN minute := minute +10; END_IF;
			IF bits[26] THEN minute := minute +20; END_IF;
			IF bits[27] THEN minute := minute +40; END_IF;
			IF minute > 59 OR (bits[21] XOR bits[22] XOR bits[23] XOR bits[24] XOR bits[25] XOR bits[26] XOR bits[27] XOR bits[28]) THEN error := TRUE; END_IF;

			(* decode hour *)
			word_temp := WORD#0;

			bool_temp:=bits[29];
			word_temp:=BIT_LOAD_W(word_temp,bool_temp,0);    (* word_temp.X0 := bits[29]; *)
			bool_temp:=bits[30];
			word_temp:=BIT_LOAD_W(word_temp,bool_temp,1);    (* word_temp.X1 := bits[30]; *)
			bool_temp:=bits[31];
			word_temp:=BIT_LOAD_W(word_temp,bool_temp,2);    (* word_temp.X2 := bits[31]; *)
			bool_temp:=bits[32];
			word_temp:=BIT_LOAD_W(word_temp,bool_temp,3);    (* word_temp.X3 := bits[32]; *)

			hour := WORD_TO_INT(word_temp);
			IF bits[33] THEN hour := hour +10; END_IF;
			IF bits[34] THEN hour := hour +20; END_IF;
			IF hour > 23 OR (bits[29] XOR bits[30] XOR bits[31] XOR bits[32] XOR bits[33] XOR bits[34] XOR bits[35]) THEN error := TRUE; END_IF;

			(* decode day of month *)
			word_temp := WORD#0;

			bool_temp:=bits[36];
			word_temp:=BIT_LOAD_W(word_temp,bool_temp,0);    (* word_temp.X0 := bits[36]; *)
			bool_temp:=bits[37];
			word_temp:=BIT_LOAD_W(word_temp,bool_temp,1);    (* word_temp.X1 := bits[37]; *)
			bool_temp:=bits[38];
			word_temp:=BIT_LOAD_W(word_temp,bool_temp,2);    (* word_temp.X2 := bits[38]; *)
			bool_temp:=bits[39];
			word_temp:=BIT_LOAD_W(word_temp,bool_temp,3);    (* word_temp.X3 := bits[39]; *)

			day := WORD_TO_INT(word_temp);
			IF bits[40] THEN day := day + 10; END_IF;
			IF bits[41] THEN day := day + 20; END_IF;
			IF day > 31 THEN error := TRUE; END_IF;

			(* decode day of week *)
			word_temp := WORD#0;

			bool_temp:=bits[42];
			word_temp:=BIT_LOAD_W(word_temp,bool_temp,0);    (* word_temp.X0 := bits[42]; *)
			bool_temp:=bits[43];
			word_temp:=BIT_LOAD_W(word_temp,bool_temp,1);    (* word_temp.X1 := bits[43]; *)
			bool_temp:=bits[44];
			word_temp:=BIT_LOAD_W(word_temp,bool_temp,2);    (* word_temp.X2 := bits[44]; *)

			wday := WORD_TO_INT(word_temp);
			IF wday > 7 OR wday < 1 THEN error := TRUE; END_IF;

			(* decode month *)
			word_temp := WORD#0;

			bool_temp:=bits[45];
			word_temp:=BIT_LOAD_W(word_temp,bool_temp,0);    (* word_temp.X0 := bits[45]; *)
			bool_temp:=bits[46];
			word_temp:=BIT_LOAD_W(word_temp,bool_temp,1);    (* word_temp.X1 := bits[46]; *)
			bool_temp:=bits[47];
			word_temp:=BIT_LOAD_W(word_temp,bool_temp,2);    (* word_temp.X2 := bits[47]; *)
			bool_temp:=bits[48];
			word_temp:=BIT_LOAD_W(word_temp,bool_temp,3);    (* word_temp.X3 := bits[48]; *)

			month := WORD_TO_INT(word_temp);
			IF bits[49] THEN month := month +10; END_IF;
			IF month > 12 THEN error := TRUE; END_IF;

			(* decode year *)
			word_temp := WORD#0;

			bool_temp:=bits[50];
			word_temp:=BIT_LOAD_W(word_temp,bool_temp,0);    (* word_temp.X0 := bits[50]; *)
			bool_temp:=bits[51];
			word_temp:=BIT_LOAD_W(word_temp,bool_temp,1);    (* word_temp.X1 := bits[51]; *)
			bool_temp:=bits[52];
			word_temp:=BIT_LOAD_W(word_temp,bool_temp,2);    (* word_temp.X2 := bits[52]; *)
			bool_temp:=bits[53];
			word_temp:=BIT_LOAD_W(word_temp,bool_temp,3);    (* word_temp.X3 := bits[53]; *)

			year := WORD_TO_INT(word_temp);
			IF bits[54] THEN year := year + 10; END_IF;
			IF bits[55] THEN year := year + 20; END_IF;
			IF bits[56] THEN year := year + 40; END_IF;
			IF bits[57] THEN year := year + 80; END_IF;

			(* check parity for bits 36 to 58 *)
			cnt := 0;
			FOR i := 36 TO 58 DO IF bits[i] THEN cnt := cnt + 1; END_IF; END_FOR;
			IF NOT even(INT_TO_DINT(cnt)) THEN error := TRUE; END_IF;

			(* time must be valid for two cycles to clear error flag *)
			IF NOT error THEN
				(* set outputs *)
				old_time := mez;
				IF year >= 70 THEN year := year + 1900; ELSE year := year + 2000; END_IF;
				mez := set_DT(year,month,day,hour,minute,0);
				DS := bits[17];
				IF DS THEN
					UTC := mez - UDINT#7200;
				ELSE
					UTC := mez - UDINT#3600;
				END_IF;

				(* set trigger signal only if the receiver has received 2 successive minutes *)
				IF mez <> old_time + TIME_TO_UDINT(t#1m) THEN error := TRUE ; END_IF;
			END_IF;
		END_IF;
	END_IF;

	tz := UDINT_TO_TIME(_INT_TO_UDINT(ABS(time_offset))* UDINT#3600000);

	IF NOT init OR SET THEN
		init := TRUE;
		utc := sdt;
		tpp := TRUE;
		DS := DSI;
	END_IF;

	IF tpp THEN
		rtc2 := utc;
		IF DS AND dst_en THEN
			IF time_offset < 0 THEN
				rtc21 := rtc2 - TIME_TO_UDINT(tz + t#1h);
			ELSE
				rtc21 := rtc2 + TIME_TO_UDINT(tz + t#1h);
			END_IF;
		ELSE
			IF time_offset < 0 THEN
				rtc21 := rtc2 - TIME_TO_UDINT(tz);
			ELSE
				rtc21 := rtc2 + TIME_TO_UDINT(tz);
			END_IF;
		END_IF;
		sync := TRUE;
		last_sync := last;
		ty := last;
	ELSIF rtc2 > UDINT#0 AND T1 - ty >= t#1s THEN
		rtc2 := rtc2 + TIME_TO_UDINT(t#1s);
		rtc21 := rtc21 + TIME_TO_UDINT(t#1s);
		ty := ty + t#1s;
		sync := ty - last_sync < sync_timeout AND last_sync > t#0s;
		wday := DAY_OF_WEEK(DT_TO_DATE2(rtc21));
		DS := dst_en AND DST(utc);
	END_IF;
	msec := TIME_TO_INT(t1 - ty);

END_FUNCTION_BLOCK

PROGRAM program0
  VAR
	REC         :	BOOL;
	SET         :	BOOL;
	SDT         :	UDINT;
	DSI         :	BOOL;
	SYNC_TIMEOUT:	TIME;
	TIME_OFFSET :	INT;
	DST_EN 	    :	BOOL;

	TPp   :	BOOL;
	DS   :	BOOL;
	WDAY :	INT;
	ERROR:	BOOL;
	RTC2  :	UDINT;
	RTC21 :	UDINT;
	MSEC :	INT;
	SYNC :	BOOL;

	func_block : DCF77;
  END_VAR
	func_block.REC           :=REC         ;
	func_block.SET           :=SET         ;
	func_block.SDT           :=SDT         ;
	func_block.DSI           :=DSI         ;
	func_block.SYNC_TIMEOUT  :=SYNC_TIMEOUT;
	func_block.TIME_OFFSET   :=TIME_OFFSET ;
	func_block.DST_EN 	      :=DST_EN 	    ;
	func_block();
	TPp   := func_block.TPp   ;
	DS   := func_block.DS   ;
	WDAY := func_block.WDAY ;
	ERROR:= func_block.ERROR;
	RTC2  := func_block.RTC2  ;
	RTC21 := func_block.RTC21 ;
	MSEC := func_block.MSEC ;
	SYNC := func_block.SYNC ;
END_PROGRAM

CONFIGURATION Config0
	VAR_GLOBAL
		PLC_TICKS_PER_SEC :	INT;
		PLC_SYS_TICK_CNT :	DINT;
	END_VAR

  	RESOURCE Res0 ON PLC
    	TASK task0(INTERVAL := T#20ms,PRIORITY := 0);
    	PROGRAM instance0 WITH task0 : program0;
  	END_RESOURCE
END_CONFIGURATION

(* ---- 735-TN_SEND_ROWS.ST ---- *)
TYPE
  oscat_IP_FIFO128_DATA  : ARRAY [1..128] OF BYTE;
  oscat_Mailbox  : ARRAY [1..16] OF BYTE;

  oscat_IP_FIFO_DATA :
  STRUCT
    X       : oscat_IP_FIFO128_DATA; (* IP_ID FIFO Speicher          *)
    Y       : oscat_IP_FIFO128_DATA; (* IP_ID Z�hler                 *)
    ID      : BYTE;                  (* h�chste vergabene id         *)
    MAX_ID  : BYTE;                  (* maximal Anmeldungen pro ID   *)
    INIT    : BOOL;                  (* Initialisierung durchgef�hrt *)
    EMPTY   : BOOL;                  (* FIFO leer                    *)
    FULL    : BOOL;                  (* FIFO voll                    *)
    TOP     : INT;                   (* maximale anzahl in FIFO      *)
    NW      : INT;                   (* Schreibzeiger                *)
    NR      : INT;                   (* Lesezeiger                   *)
  END_STRUCT;

  oscat_IP_C:
  STRUCT
    C_MODE:			BYTE;          		(*W Mode: TCP/UCP AKTIV/PASSIV                               *)
    C_PORT:         WORD;          		(*W Portnummer                                               *)
    C_IP:           DWORD;         		(*W IP-Adresse gepackt wwxxyyzz = www.xxx.yyy.zzz            *)
    C_STATE:        BYTE;          		(*R Verbindungsstatus ON/OFF + Flanke ON/OFF                 *)
    C_ENABLE:       BOOL;          		(*W Freigabe f�r Connect                                     *)
    R_OBSERVE:      BOOL;          		(*W Empfang ueberwachen                                      *)
    TIME_RESET:     BOOL;          		(*W Alle Timer ruecksetzen                                   *)
    ERROR:          DWORD;         		(*R vvwwxxyy (vv = CON_ERROR, ww = SEN_ERROR, xx = REC_ERROR *)
    FIFO:           oscat_IP_FIFO_DATA; (*I IP FIFO Struktur                                         *)
    MAILBOX:		oscat_Mailbox;		(*I Mailbox: Datenbereich f�r Bausteindatenaustausch         *)
    END_STRUCT;
END_TYPE

TYPE

  oscat_NW_BUF_LONG  : ARRAY [0..4095] OF BYTE;

  oscat_NETWORK_BUFFER :
  STRUCT
    SIZE   : UINT;
    BUFFER : oscat_NW_BUF_LONG;
  END_STRUCT;

END_TYPE

TYPE

  bya_TN_CHAR:       	ARRAY [0..1919] OF BYTE;
  bya_TN_BACKUP:     	ARRAY [0..1919] OF BYTE;
  bya_TN_COLOR:      	ARRAY [0..1919] OF BYTE;
  bya_TN_Line_Update:	ARRAY [0..23]   OF BOOL;

  us_TN_SCREEN :
  STRUCT
    bya_CHAR:			bya_TN_CHAR;
    bya_COLOR:			bya_TN_COLOR;
    bya_BACKUP:			bya_TN_BACKUP;
    bya_Line_Update:	bya_TN_Line_Update;

    by_Input_Exten_Code:    BYTE;
    by_Input_ASCII_Code:    BYTE;
    bo_Input_ASCII_IsNum:   BOOL;
    in_Page_Number:        	INT;                (* aktive Seiten-Nr.              *)
    in_Cursor_X:           	INT;                (* Cursor X-Position              *)
    in_Cursor_Y:           	INT;                (* Cursor Y-Position              *)
    in_EOS_Offset:         	INT;                (* End of String Offset           *)
    by_Clear_Screen_Attr:  	BYTE;               (* Clear-Screen Attr              *)
    bo_Clear_Screen:       	BOOL;               (* Clear-Screen ausl�sen          *)
    bo_Modal_Dialog:       	BOOL;               (* Modaler Dialog ist aktiv       *)
    bo_Menue_Bar_Dialog:   	BOOL;               (* Menue Dialog ist aktiv         *)

  END_STRUCT;
END_TYPE

FUNCTION INT_TO_BCDC:BYTE

	VAR_INPUT
		IN :	INT;
	END_VAR

	INT_TO_BCDC := SHL(INT_TO_BYTE(IN / INT#10),4) OR INT_TO_BYTE(in MOD INT#10);

END_FUNCTION

FUNCTION_BLOCK TN_SEND_ROWS_Block

  VAR_IN_OUT
    IP_C :	oscat_IP_C;
    S_BUF :	oscat_NETWORK_BUFFER;
    Xus_TN_SCREEN :	us_TN_SCREEN;
  END_VAR

  VAR_INPUT
    S_BUF_SIZE :	INT;
  END_VAR

  VAR
    in_Line_Count :	INT;
    in_Col_Count :	INT;
    in_Last_Row_Index :	INT;
    bo_Break_Loop :	BOOL;
    in_Row_Count :	INT;
    in_Offset :	INT;
    in_Write_Index :	INT;
    in_Write_Index_Backup :	INT;
    by_Cur_Color :	BYTE;
    by_last_Color :	BYTE;
    in_Write_Stop :	INT;
  END_VAR

  IF (IP_C.C_STATE < BYTE#127 OR S_BUF.SIZE > UINT#0) THEN
    RETURN;
  END_IF;

  in_Write_Index := UINT_TO_INT(S_BUF.SIZE) - 1;

  in_Write_Index_Backup := in_Write_Index;

  IF (IP_C.C_STATE = BYTE#254) OR (Xus_TN_SCREEN.bo_Clear_Screen) THEN

    Xus_TN_SCREEN.bo_Clear_Screen := FALSE;

    FOR in_Line_Count := INT#00 TO INT#23 DO
      Xus_TN_SCREEN.bya_Line_Update[in_Line_Count] := TRUE;
    END_FOR;

    in_Write_Index := in_Write_Index + INT#1;
    S_BUF.BUFFER[in_Write_Index] := BYTE#16#1B;
    in_Write_Index := in_Write_Index + INT#1;
    S_BUF.BUFFER[in_Write_Index] := BYTE#16#5B;
    in_Write_Index := in_Write_Index + INT#1;
    S_BUF.BUFFER[in_Write_Index] := BYTE#16#30;
    in_Write_Index := in_Write_Index + INT#1;
    S_BUF.BUFFER[in_Write_Index] := BYTE#16#3B;
    in_Write_Index := in_Write_Index + INT#1;
    S_BUF.BUFFER[in_Write_Index] := BYTE#16#33;

    in_Write_Index := in_Write_Index + INT#1;
    S_BUF.BUFFER[in_Write_Index] := (SHR(Xus_TN_SCREEN.by_Clear_Screen_Attr,4) OR BYTE#16#30);

    in_Write_Index := in_Write_Index + INT#1;
    S_BUF.BUFFER[in_Write_Index] := BYTE#16#3B;
    in_Write_Index := in_Write_Index + INT#1;
    S_BUF.BUFFER[in_Write_Index] := BYTE#16#34;

    in_Write_Index := in_Write_Index + INT#1;
    S_BUF.BUFFER[in_Write_Index] := ((Xus_TN_SCREEN.by_Clear_Screen_Attr AND BYTE#16#07) OR BYTE#16#30);

    in_Write_Index := in_Write_Index + INT#1;
    S_BUF.BUFFER[in_Write_Index] := BYTE#16#6D;

    in_Write_Index := in_Write_Index + INT#1;
    S_BUF.BUFFER[in_Write_Index] := BYTE#16#1B;
    in_Write_Index := in_Write_Index + INT#1;
    S_BUF.BUFFER[in_Write_Index] := BYTE#16#5B;
    in_Write_Index := in_Write_Index + INT#1;
    S_BUF.BUFFER[in_Write_Index] := BYTE#16#32;
    in_Write_Index := in_Write_Index + INT#1;
    S_BUF.BUFFER[in_Write_Index] := BYTE#16#4A;

    in_Write_Index := in_Write_Index + INT#1;
    S_BUF.BUFFER[in_Write_Index] := BYTE#16#1B;
    in_Write_Index := in_Write_Index + INT#1;
    S_BUF.BUFFER[in_Write_Index] := BYTE#16#5B;
    in_Write_Index := in_Write_Index + INT#1;
    S_BUF.BUFFER[in_Write_Index] := BYTE#16#3F;
    in_Write_Index := in_Write_Index + INT#1;
    S_BUF.BUFFER[in_Write_Index] := BYTE#16#37;
    in_Write_Index := in_Write_Index + INT#1;
    S_BUF.BUFFER[in_Write_Index] := BYTE#16#6C;

  END_IF;

  in_Last_Row_Index := INT#0;
  bo_Break_Loop := FALSE;
  in_Write_Stop := S_BUF_SIZE-20;

  FOR in_Line_Count := 0 TO 23 DO

    in_Offset := in_Row_Count * INT#80;

    IF (Xus_TN_SCREEN.bya_Line_Update[in_Row_Count] = TRUE) THEN

      in_Write_Index := in_Write_Index + INT#1;
      S_BUF.BUFFER[in_Write_Index] := BYTE#16#1B;
      in_Write_Index := in_Write_Index + INT#1;
      S_BUF.BUFFER[in_Write_Index] := BYTE#16#5B;

      in_Write_Index := in_Write_Index + INT#1;
      S_BUF.BUFFER[in_Write_Index] :=
        SHR(INT_TO_BCDC(in_Row_Count + INT#1),INT#4) OR BYTE#16#30;

      in_Write_Index := in_Write_Index + INT#1;
      S_BUF.BUFFER[in_Write_Index] :=
        (INT_TO_BCDC(in_Row_Count + INT#1) AND BYTE#16#0F) OR BYTE#16#30;

      in_Write_Index := in_Write_Index + INT#1;
      S_BUF.BUFFER[in_Write_Index] := BYTE#16#3B;
      in_Write_Index := in_Write_Index + INT#1;
      S_BUF.BUFFER[in_Write_Index] := BYTE#16#31;
      in_Write_Index := in_Write_Index + INT#1;
      S_BUF.BUFFER[in_Write_Index] := BYTE#16#48;

      FOR in_Col_Count := 0 TO 79 DO

        by_Cur_Color := Xus_TN_SCREEN.bya_COLOR[in_Offset];
        IF (by_Cur_Color <> by_last_Color) OR (in_Col_Count = INT#00) THEN

          in_Write_Index := in_Write_Index + INT#1;
          S_BUF.BUFFER[in_Write_Index] := BYTE#16#1B;

          in_Write_Index := in_Write_Index + INT#1;
          S_BUF.BUFFER[in_Write_Index] := BYTE#16#5B;

          IF  (((by_Cur_Color AND BYTE#2#10001000) XOR (by_last_Color AND BYTE#2#10001000)) <> BYTE#00) OR (in_Col_Count = 0) THEN

            in_Write_Index := in_Write_Index + INT#1;
            S_BUF.BUFFER[in_Write_Index] := BYTE#16#30;
            in_Write_Index := in_Write_Index + INT#1;
            S_BUF.BUFFER[in_Write_Index] := BYTE#16#3B;

            IF (by_Cur_Color AND BYTE#2#00001000) = BYTE#2#00000000 THEN

              in_Write_Index := in_Write_Index + INT#1;
              S_BUF.BUFFER[in_Write_Index] := BYTE#16#31;
              in_Write_Index := in_Write_Index + INT#1;
              S_BUF.BUFFER[in_Write_Index] := BYTE#16#3B;

            END_IF;

            IF (by_Cur_Color AND BYTE#2#10000000) = BYTE#2#10000000 THEN

              in_Write_Index := in_Write_Index + INT#1;
              S_BUF.BUFFER[in_Write_Index] := BYTE#16#35;
              in_Write_Index := in_Write_Index + INT#1;
              S_BUF.BUFFER[in_Write_Index] := BYTE#16#3B;

            END_IF;

          END_IF;

          in_Write_Index := in_Write_Index + INT#1;
          S_BUF.BUFFER[in_Write_Index] := BYTE#16#33;

          in_Write_Index := in_Write_Index + INT#1;
          S_BUF.BUFFER[in_Write_Index] := ((SHR(by_Cur_Color,4) AND BYTE#2#00000111) OR BYTE#16#30);

          in_Write_Index := in_Write_Index + INT#1;
          S_BUF.BUFFER[in_Write_Index] := BYTE#16#3B;

          in_Write_Index := in_Write_Index + INT#1;
          S_BUF.BUFFER[in_Write_Index] := BYTE#16#34;

          in_Write_Index := in_Write_Index + INT#1;
          S_BUF.BUFFER[in_Write_Index] := ((by_Cur_Color AND BYTE#2#00000111) OR BYTE#16#30);

          in_Write_Index := in_Write_Index + INT#1;
          S_BUF.BUFFER[in_Write_Index] := BYTE#16#6D;

          by_last_Color := by_Cur_Color;

        END_IF;

        IF (in_Write_Index > in_Write_Stop) THEN

          bo_Break_Loop := TRUE;
          EXIT;

        END_IF;

        in_Write_Index := in_Write_Index + INT#1;
        S_BUF.BUFFER[in_Write_Index] := Xus_TN_SCREEN.bya_CHAR[in_Offset];

        in_Offset := in_Offset + INT#01;
      END_FOR;

      IF (bo_Break_Loop = TRUE) THEN

        in_Write_Index := in_Last_Row_Index;

        EXIT;
      END_IF;

      in_Last_Row_Index := in_Write_Index;
      Xus_TN_SCREEN.bya_Line_Update[in_Row_Count] := FALSE;

    END_IF;

    in_Row_Count := in_Row_Count + INT#01;

    IF (in_Row_Count > INT#23) THEN
      in_Row_Count := INT#00;
    END_IF;

  END_FOR;

  IF (bo_Break_Loop = FALSE) THEN

    in_Row_Count := INT#00;

  END_IF;

  IF (in_Write_Index <> in_Write_Index_Backup) THEN

    in_Write_Index := in_Write_Index + INT#1;
    S_BUF.BUFFER[in_Write_Index] := BYTE#16#1B;
    in_Write_Index := in_Write_Index + INT#1;
    S_BUF.BUFFER[in_Write_Index] := BYTE#16#5B;

    in_Write_Index := in_Write_Index + INT#1;
    S_BUF.BUFFER[in_Write_Index] := SHR(INT_TO_BCDC(Xus_TN_SCREEN.in_Cursor_Y + 1),INT#4) OR BYTE#16#30;

    in_Write_Index := in_Write_Index + INT#1;
    S_BUF.BUFFER[in_Write_Index] := (INT_TO_BCDC(Xus_TN_SCREEN.in_Cursor_Y + 1) AND BYTE#16#0F) OR BYTE#16#30;

    in_Write_Index := in_Write_Index + INT#1;
    S_BUF.BUFFER[in_Write_Index] := BYTE#16#3B;

    in_Write_Index := in_Write_Index + INT#1;
    S_BUF.BUFFER[in_Write_Index] := SHR(INT_TO_BCDC(Xus_TN_SCREEN.in_Cursor_X + 1),INT#4) OR BYTE#16#30;

    in_Write_Index := in_Write_Index + INT#1;
    S_BUF.BUFFER[in_Write_Index] := (INT_TO_BCDC(Xus_TN_SCREEN.in_Cursor_X + 1) AND BYTE#16#0F) OR BYTE#16#30;

    in_Write_Index := in_Write_Index + INT#1;
    S_BUF.BUFFER[in_Write_Index] := BYTE#16#48;

  END_IF;

  S_BUF.SIZE := INT_TO_UINT(in_Write_Index + 1);

END_FUNCTION_BLOCK

PROGRAM program0
	VAR
		IP_C :	oscat_IP_C;
    S_BUF :	oscat_NETWORK_BUFFER;
    Xus_TN_SCREEN :	us_TN_SCREEN;
    S_BUF_SIZE :	INT;

		func_block : TN_SEND_ROWS_Block;
	END_VAR
	func_block.IP_C := IP_C;
  func_block.S_BUF := S_BUF;
  func_block.Xus_TN_SCREEN := Xus_TN_SCREEN;
  func_block.S_BUF_SIZE := S_BUF_SIZE;

	func_block();
	IP_C  := func_block.IP_C;
  S_BUF  := func_block.S_BUF;
  Xus_TN_SCREEN  := func_block.Xus_TN_SCREEN;
END_PROGRAM

CONFIGURATION Config0
	RESOURCE Res0 ON PLC
		TASK task0(INTERVAL := T#20ms,PRIORITY := 0);
		PROGRAM instance0 WITH task0 : program0;
	END_RESOURCE
END_CONFIGURATION

(* ---- 736-TEMP_EXT.ST ---- *)
FUNCTION UDINT_TO_TIME2:TIME

	VAR_INPUT
		IN :	UDINT;
	END_VAR

	UDINT_TO_TIME2 := DINT_TO_TIME(UDINT_TO_DINT(IN));

END_FUNCTION

FUNCTION_BLOCK T_PLC_MS_block
	VAR_OUTPUT
		T_PLC_MS :	UDINT;
	END_VAR

	VAR_EXTERNAL
		PLC_TICKS_PER_SEC :	INT;
		PLC_SYS_TICK_CNT :	DINT;
	END_VAR

	VAR
		debug :	BOOL;(*Debug-Mode ON / OFF*)
		N :	INT;(*Debug-Faktor*)
		Offset :	UDINT;(*Debug-Offset*)
		temp :	DWORD := DWORD#1;(*Debug-Offset*)
		mode :	BOOL;(*modus*)
		faktor :	UDINT;(*Systemtakt-Faktor*)
		init :	BOOL;
		v_plc_ticks_per_sec :	UDINT;
		base :	UDINT := UDINT#1000;
	END_VAR

	IF init = FALSE THEN
		v_plc_ticks_per_sec := INT_TO_UDINT(PLC_TICKS_PER_SEC);
		IF v_plc_ticks_per_sec = UDINT#1024 THEN
			faktor := UDINT#1;
			mode := FALSE;
		ELSIF v_plc_ticks_per_sec > UDINT#0 THEN
			IF v_plc_ticks_per_sec <= base THEN
				faktor := base / v_plc_ticks_per_sec;
				mode := FALSE;
			ELSE
				faktor := v_plc_ticks_per_sec / base;
				mode := TRUE;
			END_IF;
		ELSE
			faktor := UDINT#1;
		END_IF;
		init := TRUE;
	END_IF;

	IF mode THEN
		T_PLC_MS := DINT_TO_UDINT(PLC_SYS_TICK_CNT) / faktor;
	ELSE
		T_PLC_MS := DINT_TO_UDINT(PLC_SYS_TICK_CNT) * faktor;
	END_IF;

	IF debug THEN
		T_PLC_MS := (DWORD_TO_UDINT(SHL(UDINT_TO_DWORD(T_PLC_MS),N) OR SHL(temp,N)) - UDINT#1) + Offset;
	END_IF;
END_FUNCTION_BLOCK

FUNCTION _INT_TO_UDINT:UDINT
	VAR_INPUT
		IN :	INT;
	END_VAR

	_INT_TO_UDINT := DINT_TO_UDINT(INT_TO_DINT(IN));
END_FUNCTION

FUNCTION SET_DATE:UDINT

	VAR_INPUT
		YEAR :	INT;
		MONTH :	INT;
		DAY :	INT;
	END_VAR

	VAR
		count :	INT;
	END_VAR

	IF month > 2 THEN
		count := (month - 1) * 30;
		IF month > 7 THEN
			count := count + DWORD_TO_INT(SHR(DINT_TO_DWORD(INT_TO_DINT(month) - INT_TO_DINT(3)),1));
		ELSE
			count := count + DWORD_TO_INT(SHR(DINT_TO_DWORD(INT_TO_DINT(month) - INT_TO_DINT(4)),1));
		END_IF;
		IF SHL(INT_TO_WORD(year),14) = WORD#0 THEN
			count := count + 1;
		END_IF;
	ELSE
		count := (month - 1) * 31;
	END_IF;
	SET_DATE := (_INT_TO_UDINT(count + day - 1) + DWORD_TO_UDINT(SHR(UDINT_TO_DWORD(_INT_TO_UDINT(year) * UDINT#1461 - UDINT#2878169), 2))) * UDINT#86400;

END_FUNCTION

FUNCTION LEAP_OF_DATE:BOOL

	VAR_INPUT
		IDATE :	UDINT;
	END_VAR

	LEAP_OF_DATE := SHL(UDINT_TO_DWORD((idate + UDINT#43200) / UDINT#31557600), 30) = DWORD#16#80000000;

END_FUNCTION

FUNCTION DAY_OF_YEAR:INT
	VAR_INPUT
		IDATE :	DATE;
	END_VAR

	DAY_OF_YEAR := UDINT_TO_INT((DATE_TO_UDINT(idate) / UDINT#86400) MOD UDINT#1461);
	IF DAY_OF_YEAR > 729 THEN
		IF DAY_OF_YEAR > 1095 THEN DAY_OF_YEAR := DAY_OF_YEAR - 1095; ELSE DAY_OF_YEAR := DAY_OF_YEAR - 729; END_IF;
	ELSIF DAY_OF_YEAR > 364 THEN
		DAY_OF_YEAR := DAY_OF_YEAR - 364;
	ELSE
		DAY_OF_YEAR := DAY_OF_YEAR + 1;
	END_IF;
END_FUNCTION

FUNCTION DAY_OF_YEAR_UDINT:INT
	VAR_INPUT
		IDATE :	UDINT;
	END_VAR

	DAY_OF_YEAR_UDINT := UDINT_TO_INT((idate / UDINT#86400) MOD UDINT#1461);
	IF DAY_OF_YEAR_UDINT > 729 THEN
		IF DAY_OF_YEAR_UDINT > 1095 THEN DAY_OF_YEAR_UDINT := DAY_OF_YEAR_UDINT - 1095; ELSE DAY_OF_YEAR_UDINT := DAY_OF_YEAR_UDINT - 729; END_IF;
	ELSIF DAY_OF_YEAR_UDINT > 364 THEN
		DAY_OF_YEAR_UDINT := DAY_OF_YEAR_UDINT - 364;
	ELSE
		DAY_OF_YEAR_UDINT := DAY_OF_YEAR_UDINT + 1;
	END_IF;
END_FUNCTION

FUNCTION MONTH_OF_DATE_UDINT:INT

	VAR_INPUT
		IDATE :	UDINT;
	END_VAR

	MONTH_OF_DATE_UDINT := DAY_OF_YEAR_UDINT(idate);
	IF MONTH_OF_DATE_UDINT < 32 THEN
		MONTH_OF_DATE_UDINT := 1;
	ELSIF LEAP_OF_DATE(IDATE) THEN
		MONTH_OF_DATE_UDINT := (MONTH_OF_DATE_UDINT * 53 + 1668) / 1623;
	ELSE
		MONTH_OF_DATE_UDINT := (MONTH_OF_DATE_UDINT * 53 + 1700) / 1620;
	END_IF;

END_FUNCTION

FUNCTION DAY_OF_MONTH:INT
	VAR_INPUT
		IDATE :	UDINT;
	END_VAR

	day_of_month := day_of_year_UDINT(idate);

	IF leap_of_Date(idate) THEN
		CASE day_of_month OF
			32..60	:	day_of_month := day_of_month - 31;
			61..91	:	day_of_month := day_of_month - 60;
			92..121 :	day_of_month := day_of_month - 91;
			122..152:	day_of_month := day_of_month - 121;
			153..182:	day_of_month := day_of_month - 152;
			183..213:	day_of_month := day_of_month - 182;
			214..244:	day_of_month := day_of_month - 213;
			245..274:	day_of_month := day_of_month - 244;
			275..305:	day_of_month := day_of_month - 274;
			306..335:	day_of_month := day_of_month - 305;
			336..366:	day_of_month := day_of_month - 335;
		END_CASE;
	ELSE
		CASE day_of_month OF
			32..59	:	day_of_month := day_of_month - 31;
			60..90	:	day_of_month := day_of_month - 59;
			91..120 :	day_of_month := day_of_month - 90;
			121..151:	day_of_month := day_of_month - 120;
			152..181:	day_of_month := day_of_month - 151;
			182..212:	day_of_month := day_of_month - 181;
			213..243:	day_of_month := day_of_month - 212;
			244..273:	day_of_month := day_of_month - 243;
			274..304:	day_of_month := day_of_month - 273;
			305..334:	day_of_month := day_of_month - 304;
			335..365:	day_of_month := day_of_month - 334;
		END_CASE;
	END_IF;

END_FUNCTION

FUNCTION MID3:REAL

	VAR_INPUT
		IN1 :	REAL;
		IN2 :	REAL;
		IN3 :	REAL;
	END_VAR

	VAR
		_IN1 :	REAL;
		_IN2 :	REAL;
		_IN3 :	REAL;
	END_VAR

	_IN1 := IN1;
	_IN2 := IN2;
	_IN3 := IN3;

	IF _IN1 > _IN2 THEN MID3 := _IN1; _IN1 := _IN2; _IN2 := MID3; END_IF;
	IF _IN2 > _IN3 THEN _IN2 := _IN3; END_IF;
	MID3 := SEL(_IN1 > _IN2, _IN2, _IN1);

END_FUNCTION

FUNCTION _BYTE_TO_INT:INT
	VAR_INPUT
		IN :	BYTE;
	END_VAR

	_BYTE_TO_INT := USINT_TO_INT(BYTE_TO_USINT(IN));
END_FUNCTION

FUNCTION MULTI_IN:REAL

	VAR_INPUT
		IN_1 :	REAL;
		IN_2 :	REAL;
		IN_3 :	REAL;
		DEFAULT :	REAL;
		IN_MIN :	REAL;
		IN_MAX :	REAL;
		MODE :	BYTE;
	END_VAR

	VAR
		count :	INT;
		F1 :	BOOL;
		F2 :	BOOL;
		F3 :	BOOL;
	END_VAR

	F1 :=  in_1 > in_min AND in_1 < in_max;
	F2 :=  in_2 > in_min AND in_2 < in_max;
	F3 :=  in_3 > in_min AND in_3 < in_max;

	CASE _BYTE_TO_INT(mode) OF
	0:	count := 0;
		IF F1 THEN
			count := count + 1;
			MULTI_IN := in_1;
		ELSE
			MULTI_IN := 0.0;
		END_IF;
		IF F2 THEN
			count := count + 1;
			MULTI_IN := MULTI_IN + in_2;
		END_IF;
		IF F3 THEN
			count := count + 1;
			MULTI_IN := MULTI_IN + in_3;
		END_IF;
		MULTI_IN := SEL_REAL(count = 0, MULTI_IN / INT_TO_REAL(count), default);

	1:	MULTI_IN := SEL_REAL(F1, default, IN_1);

	2:	MULTI_IN := SEL_REAL(F2, default, IN_2);

	3:	MULTI_IN := SEL_REAL(F3, default, IN_3);

	4:	MULTI_IN := default;

	5:	MULTI_IN := SEL_REAL(F1, in_max, IN_1);
		IF F2 AND in_2 < MULTI_IN THEN MULTI_IN := in_2; END_IF;
		IF F3 AND in_3 < MULTI_IN THEN MULTI_IN := in_3; END_IF;
		IF MULTI_IN = in_max THEN MULTI_IN := default; END_IF;

	6:	MULTI_IN := SEL_REAL(F1, in_min, IN_1);
		IF F2 AND in_2 > MULTI_IN THEN MULTI_IN := in_2; END_IF;
		IF F3 AND in_3 > MULTI_IN THEN MULTI_IN := in_3; END_IF;
		IF MULTI_IN = in_min THEN MULTI_IN := default; END_IF;

	7:	IF F1 AND F2 AND F3 THEN MULTI_IN := MID3(in_1, in_2, in_3);
		ELSIF F1 AND F2 THEN MULTI_IN := MIN(in_1, in_2);
		ELSIF F1 AND F3 THEN MULTI_IN := MIN(in_1, in_3);
		ELSIF F2 AND F3 THEN MULTI_IN := MIN(in_2, in_3);
		ELSIF F1 THEN MULTI_IN := in_1;
		ELSIF F2 THEN MULTI_IN := in_2;
		ELSIF F3 THEN MULTI_IN := in_3;
		ELSE MULTI_IN := default;
		END_IF;

	END_CASE;

END_FUNCTION

FUNCTION _DT_TO_DATE_B:UDINT

	VAR_INPUT
		_INN :	UDINT;
	END_VAR

	_DT_TO_DATE_B := (_INN / UDINT#86400) * UDINT#86400;
END_FUNCTION

FUNCTION DT_TO_TOD2:UDINT
	VAR_INPUT
		IN :	UDINT;
	END_VAR

	DT_TO_TOD2 := (IN MOD UDINT#86400) * UDINT#1000;
END_FUNCTION

FUNCTION_BLOCK TEMP_EXT_Block

	VAR_INPUT
		T_EXT1 :	REAL;
		T_EXT2 :	REAL;
		T_EXT3 :	REAL;
		T_EXT_CONFIG :	BYTE := 0;
		DT_IN :	UDINT;
		T_EXT_MIN :	REAL := REAL#-40.0;
		T_EXT_MAX :	REAL := REAL#60.0;
		T_EXT_DEFAULT :	REAL := REAL#-10.0;
		HEAT_PERIOD_START :	UDINT := UDINT#20995200;
		HEAT_PERIOD_STOP :	UDINT := UDINT#10281600;
		COOL_PERIOD_START :	UDINT := UDINT#07776000;
		COOL_PERIOD_STOP :	UDINT := UDINT#23500800;
		HEAT_START_TEMP_DAY :	REAL := REAL#15.0;
		HEAT_START_TEMP_NIGHT :	REAL := REAL#10.0;
		HEAT_STOP_TEMP :	REAL := REAL#18.0;
		COOL_START_TEMP_DAY :	REAL := REAL#26.0;
		COOL_START_TEMP_NIGHT :	REAL := REAL#26.0;
		COOL_STOP_TEMP :	REAL := REAL#24.0;
		START_DAY :	UDINT := UDINT#32400000;
		START_NIGHT :	UDINT := UDINT#75600000;
		CYCLE_TIME :	TIME := t#10m;
	END_VAR

	VAR_OUTPUT
		T_EXT :	REAL;
		HEAT :	BOOL;
		COOL :	BOOL;
	END_VAR

	VAR
		tx :	TIME;
		last_run :	TIME;
		init :	BOOL;
		cool_start :	UDINT;
		cool_stop :	UDINT;
		heat_start :	UDINT;
		heat_stop :	UDINT;
		xdate :	UDINT;
		day :	BOOL;
		T_PLC_MS :	T_PLC_MS_Block;
	END_VAR

	IF NOT init THEN
		init := TRUE;
		heat_start := SET_DATE(1972,MONTH_OF_DATE_UDINT(heat_period_start),DAY_OF_MONTH(heat_period_start));
		heat_stop := SET_DATE(1972,MONTH_OF_DATE_UDINT(heat_period_stop),DAY_OF_MONTH(heat_period_stop));
		cool_start := SET_DATE(1972,MONTH_OF_DATE_UDINT(cool_period_start),DAY_OF_MONTH(cool_period_start));
		cool_stop := SET_DATE(1972,MONTH_OF_DATE_UDINT(cool_period_stop),DAY_OF_MONTH(cool_period_stop));
	END_IF;

	T_PLC_MS();
	tx:= UDINT_TO_TIME(T_PLC_MS.T_PLC_MS);

	IF tx - last_run < cycle_time THEN RETURN; END_IF;

	xdate := SET_DATE(1972,MONTH_OF_DATE_UDINT(_DT_TO_DATE_B(dt_in)),DAY_OF_MONTH(_DT_TO_DATE_B(dt_in)));
	day := DT_TO_TOD2(dt_in) >= start_day AND  DT_TO_TOD2(dt_in) < start_night;

	t_ext := MULTI_IN(t_ext1, t_ext2, t_ext3, t_ext_default, t_ext_min, t_ext_max, t_ext_config);

	IF (heat_start <= heat_stop AND xdate >= heat_start AND xdate <= heat_stop) OR (heat_start > heat_stop AND (xdate >= heat_start OR xdate <= heat_stop)) THEN
		IF day AND t_ext <= heat_start_temp_day THEN
			heat := TRUE;
		ELSIF NOT day AND t_ext <= heat_start_temp_night THEN
			heat := TRUE;
		ELSIF t_ext >= heat_stop_temp THEN
			heat := FALSE;
		END_IF;
	ELSE
		heat := FALSE;
	END_IF;

	IF (cool_start <= cool_stop AND xdate >= cool_start AND xdate <= cool_stop) OR (cool_start > cool_stop AND (xdate >= cool_start OR xdate <= cool_stop)) THEN
		IF day AND t_ext >= cool_start_temp_day THEN
			cool := TRUE;
		ELSIF NOT day AND t_ext >= cool_start_temp_night THEN
			cool := TRUE;
		ELSIF t_ext <= cool_stop_temp THEN
			cool := FALSE;
		END_IF;
	ELSE
		cool := FALSE;
	END_IF;

	last_run := tx;

END_FUNCTION_BLOCK

PROGRAM program0
	VAR
		T_EXT1 :	REAL;
		T_EXT2 :	REAL;
		T_EXT3 :	REAL;
		T_EXT_CONFIG :	BYTE := 0;
		DT_IN :	UDINT;
		T_EXT_MIN :	REAL := REAL#-40.0;
		T_EXT_MAX :	REAL := REAL#60.0;
		T_EXT_DEFAULT :	REAL := REAL#-10.0;
		HEAT_PERIOD_START :	UDINT := UDINT#20995200;
		HEAT_PERIOD_STOP :	UDINT := UDINT#10281600;
		COOL_PERIOD_START :	UDINT := UDINT#07776000;
		COOL_PERIOD_STOP :	UDINT := UDINT#23500800;
		HEAT_START_TEMP_DAY :	REAL := REAL#15.0;
		HEAT_START_TEMP_NIGHT :	REAL := REAL#10.0;
		HEAT_STOP_TEMP :	REAL := REAL#18.0;
		COOL_START_TEMP_DAY :	REAL := REAL#26.0;
		COOL_START_TEMP_NIGHT :	REAL := REAL#26.0;
		COOL_STOP_TEMP :	REAL := REAL#24.0;
		START_DAY :	UDINT := UDINT#32400000;
		START_NIGHT :	UDINT := UDINT#75600000;
		CYCLE_TIME :	TIME := t#10m;
		T_EXT :	REAL;
		HEAT :	BOOL;
		COOL :	BOOL;

		func_block : TEMP_EXT_Block;
	END_VAR

	func_block.T_EXT1 := T_EXT1;
	func_block.T_EXT2 := T_EXT2;
	func_block.T_EXT3 := T_EXT3 ;
	func_block.T_EXT_CONFIG := T_EXT_CONFIG;
	func_block.DT_IN := DT_IN;
	func_block.T_EXT_MIN := T_EXT_MIN ;
	func_block.T_EXT_MAX := T_EXT_MAX;
	func_block.T_EXT_DEFAULT := T_EXT_DEFAULT;
	func_block.HEAT_PERIOD_START := HEAT_PERIOD_START ;
	func_block.HEAT_PERIOD_STOP := HEAT_PERIOD_STOP;
	func_block.COOL_PERIOD_START := COOL_PERIOD_START;
	func_block.COOL_PERIOD_STOP := COOL_PERIOD_STOP ;
	func_block.HEAT_START_TEMP_DAY := HEAT_START_TEMP_DAY;
	func_block.HEAT_START_TEMP_NIGHT := HEAT_START_TEMP_NIGHT;
	func_block.HEAT_STOP_TEMP := HEAT_STOP_TEMP ;
	func_block.COOL_START_TEMP_DAY := COOL_START_TEMP_DAY;
	func_block.COOL_START_TEMP_NIGHT := COOL_START_TEMP_NIGHT;
	func_block.COOL_STOP_TEMP:= COOL_STOP_TEMP ;
	func_block.START_DAY := START_DAY;
	func_block.START_NIGHT := START_NIGHT;
	func_block.CYCLE_TIME:= CYCLE_TIME ;

	func_block();
	T_EXT  := func_block.T_EXT;
	HEAT  := func_block.HEAT;
	COOL  := func_block.COOL;

END_PROGRAM

CONFIGURATION Config0
	VAR_GLOBAL
		PLC_TICKS_PER_SEC :	INT;
		PLC_SYS_TICK_CNT :	DINT;
	END_VAR
  	RESOURCE Res0 ON PLC
    	TASK task0(INTERVAL := T#20ms,PRIORITY := 0);
    	PROGRAM instance0 WITH task0 : program0;
  	END_RESOURCE
END_CONFIGURATION

(* ---- 739-TELNET_PRINT.ST ---- *)
TYPE
  oscat_STRING250             : STRING;
END_TYPE

TYPE
  oscat_IP_FIFO128_DATA  : ARRAY [1..128] OF BYTE;
  oscat_Mailbox  : ARRAY [1..16] OF BYTE;

  oscat_IP_FIFO_DATA :
  STRUCT
	X       : oscat_IP_FIFO128_DATA; (* IP_ID FIFO Speicher          *)
	Y       : oscat_IP_FIFO128_DATA; (* IP_ID Z�hler                 *)
	ID      : BYTE;                  (* h�chste vergabene id         *)
	MAX_ID  : BYTE;                  (* maximal Anmeldungen pro ID   *)
    INIT    : BOOL;                  (* Initialisierung durchgef�hrt *)
	EMPTY   : BOOL;                  (* FIFO leer                    *)
	FULL    : BOOL;                  (* FIFO voll                    *)
	TOP     : INT;                   (* maximale anzahl in FIFO      *)
	NW      : INT;                   (* Schreibzeiger                *)
	NR      : INT;                   (* Lesezeiger                   *)
  END_STRUCT;

  oscat_IP_C:
  STRUCT
  	C_MODE:			BYTE;          		(*W Mode: TCP/UCP AKTIV/PASSIV                               *)
	C_PORT:         WORD;          		(*W Portnummer                                               *)
	C_IP:           DWORD;         		(*W IP-Adresse gepackt wwxxyyzz = www.xxx.yyy.zzz            *)
    C_STATE:        BYTE;          		(*R Verbindungsstatus ON/OFF + Flanke ON/OFF                 *)
	C_ENABLE:       BOOL;          		(*W Freigabe f�r Connect                                     *)
    R_OBSERVE:      BOOL;          		(*W Empfang ueberwachen                                      *)
    TIME_RESET:     BOOL;          		(*W Alle Timer ruecksetzen                                   *)
	ERROR:          DWORD;         		(*R vvwwxxyy (vv = CON_ERROR, ww = SEN_ERROR, xx = REC_ERROR *)
    FIFO:           oscat_IP_FIFO_DATA; (*I IP FIFO Struktur                                         *)
	MAILBOX:		oscat_Mailbox;		(*I Mailbox: Datenbereich f�r Bausteindatenaustausch         *)
  END_STRUCT;
END_TYPE

FUNCTION _BYTE_TO_INT:INT
	VAR_INPUT
		IN :	BYTE;
	END_VAR

	_BYTE_TO_INT := USINT_TO_INT(BYTE_TO_USINT(IN));
END_FUNCTION

FUNCTION_BLOCK IP_FIFO_Block

  VAR_IN_OUT
    FIFO :	oscat_IP_FIFO_DATA;
    ID :	BYTE;
    STATE :	BYTE;
  END_VAR

  VAR
    tmp :	INT;
  END_VAR

  IF NOT FIFO.INIT THEN
    FIFO.INIT		:= TRUE;
    FIFO.NW		:= 1;
    FIFO.NR		:= 1;
    FIFO.EMPTY	:= TRUE;
    FIFO.FULL		:= FALSE;
    FIFO.TOP		:= 128;
    FIFO.MAX_ID	:= BYTE#1;
  END_IF;

  IF ID = BYTE#00 THEN
    IF FIFO.ID < INT_TO_BYTE(FIFO.TOP) THEN
      ID := USINT_TO_BYTE(BYTE_TO_USINT(FIFO.ID) + USINT#1);
      FIFO.ID := ID ;

    ELSIF STATE < BYTE#200 THEN
      STATE := BYTE#255;
    RETURN;
    END_IF;
  END_IF;

  IF STATE = BYTE#1 AND NOT FIFO.FULL THEN
    tmp := _BYTE_TO_INT(ID);
    IF FIFO.Y[tmp] < FIFO.MAX_ID THEN
      FIFO.Y[tmp] := USINT_TO_BYTE(BYTE_TO_USINT(FIFO.Y[tmp]) + USINT#1);
      tmp := FIFO.NW;
      FIFO.X[tmp] := ID;
      IF FIFO.NW = FIFO.TOP THEN FIFO.NW := 1; ELSE FIFO.NW := FIFO.NW + 1; END_IF;
      FIFO.FULL := FIFO.NW = FIFO.NR;
    FIFO.EMPTY := FALSE;
      STATE := BYTE#2;
    END_IF;
  END_IF;

  IF STATE = BYTE#2 AND NOT FIFO.EMPTY THEN
    tmp := FIFO.NR;
    IF ID = FIFO.X[tmp] THEN
      STATE := BYTE#3;
    END_IF;
  END_IF;

  IF STATE = BYTE#4 AND NOT FIFO.EMPTY THEN

    tmp := FIFO.NR;
    IF ID = FIFO.X[tmp] THEN
      tmp := _BYTE_TO_INT(ID);
      FIFO.Y[tmp] := USINT_TO_BYTE(BYTE_TO_USINT(FIFO.Y[tmp]) - USINT#1);

      IF FIFO.NR = FIFO.TOP THEN FIFO.NR := 1; ELSE FIFO.NR := FIFO.NR + 1; END_IF;
      FIFO.EMPTY := FIFO.NR = FIFO.NW;
    FIFO.FULL := FALSE;
    END_IF;
    STATE := BYTE#5;
  END_IF;

END_FUNCTION_BLOCK

FUNCTION_BLOCK TELNET_PRINT_Block

	VAR_INPUT
		TEXT :	oscat_STRING250;
		ENABLE :	BOOL;
		SEND :	BOOL;
		OPTION :	BYTE;
		BACK_COLOR :	BYTE;
		FRONT_COLOR :	BYTE;
		X_POS :	BYTE;
		Y_POS :	BYTE;
		PORT :	WORD := WORD#23;
	END_VAR

	VAR_OUTPUT
		READY :	BOOL;
		DONE :	BOOL;
	END_VAR

	VAR_IN_OUT
		IP_C :	oscat_IP_C;
		S_BUF :	oscat_NETWORK_BUFFER;
	END_VAR

	VAR
		_STRING_TO_BUFFER :	_STRING_TO_BUFFER_NW;
		last_fc :	BYTE;
		state :	INT;
		x :	INT := -1;
		ip_state :	BYTE;
		ip_id :	BYTE;
		IP_FIFO :	IP_FIFO_Block;
		s_buf_size :	UINT := uint#4096;
		init :	BOOL;
		b0_screen_clear :	BOOL;
		b1_autowrap :	BOOL;
		b2_color :	BOOL;
		b3_cr_lr :	BOOL;
		b7_no_flush :	BOOL;
	END_VAR

	READY := IP_C.C_STATE > BYTE#127;
	DONE := FALSE;

	CASE state OF

	00:
		IF ENABLE THEN
			state := 10;
			ip_state := BYTE#1;
		END_IF;

	10:
		IF ip_state = BYTE#3 THEN

			IP_C.C_PORT := PORT;
			IP_C.C_IP := DWORD#00;
			IP_C.C_MODE := BYTE#4;
			IP_C.TIME_RESET := TRUE;
			IP_C.C_ENABLE := TRUE;
			IP_C.R_OBSERVE := FALSE;
			state := 20;
		END_IF;

	20:	IF IP_C.ERROR > DWORD#0 THEN
			IP_C.TIME_RESET := TRUE;
		END_IF;
		IF S_BUF.SIZE = UINT#0 THEN
			IF NOT ENABLE THEN
				ip_state := BYTE#4;
				IP_C.C_ENABLE := FALSE;
				state := 0;
			END_IF;
			IF IP_C.C_STATE = BYTE#1 THEN
				init := FALSE;
			ELSIF READY THEN
				IF IP_C.C_STATE = BYTE#254 AND NOT INIT THEN
					init := TRUE;
					b0_screen_clear := (OPTION AND BYTE#2#0000_0001) > BYTE#0;
					b1_autowrap := (OPTION AND BYTE#2#0000_0010) > BYTE#0;
					b2_color := (OPTION AND BYTE#2#0000_0100) > BYTE#0;
					b3_cr_lr := (OPTION AND BYTE#2#0000_1000) > BYTE#0;
					b7_no_flush := (OPTION AND BYTE#2#1000_0000) > BYTE#0;

					last_fc := NOT FRONT_COLOR;
					x := 0;

					S_BUF.BUFFER[x] := BYTE#16#1B;
					x := x +1;
					S_BUF.BUFFER[x] := BYTE#16#5B;
					x := x +1;
					S_BUF.BUFFER[x] := BYTE#16#3F;
					x := x +1;
					S_BUF.BUFFER[x] := BYTE#16#37; (
					x := x +1;
					S_BUF.BUFFER[x] := SEL(b1_autowrap, BYTE#16#6C, BYTE#16#68 );

					IF b0_screen_clear THEN
						IF b2_color THEN
							x := x +1;
							S_BUF.BUFFER[x] := BYTE#16#1B;
							x := x +1;
							S_BUF.BUFFER[x] := BYTE#16#5B;
							x := x +1;
							S_BUF.BUFFER[x] := BYTE#16#30;
							x := x +1;
							S_BUF.BUFFER[x] := BYTE#16#3B;
							x := x +1;
							S_BUF.BUFFER[x] := BYTE#16#33;
							x := x +1;
							S_BUF.BUFFER[x] := (FRONT_COLOR AND BYTE#2#00000111) OR BYTE#16#30;
							x := x +1;
							S_BUF.BUFFER[x] := BYTE#16#3B;
							x := x +1;
							S_BUF.BUFFER[x] := BYTE#16#34;
							x := x +1;
							S_BUF.BUFFER[x] := (BACK_COLOR AND BYTE#2#00000111) OR BYTE#16#30;
							x := x +1;
							S_BUF.BUFFER[x] := BYTE#16#6D;
						END_IF;
						x := x +1;
						S_BUF.BUFFER[x] := BYTE#16#1B;
						x := x +1;
						S_BUF.BUFFER[x] := BYTE#16#5B;
						x := x +1;
						S_BUF.BUFFER[x] := BYTE#16#32;
						x := x +1;
						S_BUF.BUFFER[x] := BYTE#16#4A;
					ELSE
						x := x +1;
						S_BUF.BUFFER[x] := BYTE#16#0A;
					END_IF;
				END_IF;

				IF (INT_TO_UINT(x + LEN(TEXT) + 21) > s_buf_size) OR (x >= 0 AND NOT SEND) THEN
					S_BUF.SIZE := INT_TO_UINT(x + 1);
					x := -1;
				ELSIF SEND THEN

					IF b2_color AND FRONT_COLOR <> last_FC THEN
						x := x + 1;
						S_BUF.BUFFER[x] := BYTE#16#1B;
						x := x + 1;
						S_BUF.BUFFER[x] := BYTE#16#5B;
						IF ((FRONT_COLOR AND BYTE#2#0001_1000) XOR (last_FC AND BYTE#2#0001_1000)) <> BYTE#00 OR TRUE THEN
							x := x + 1;
							S_BUF.BUFFER[x] := BYTE#16#30;
							x := x + 1;
							S_BUF.BUFFER[x] := BYTE#16#3B;
							IF (FRONT_COLOR AND BYTE#2#00001000) = BYTE#0 THEN
								x := x + 1;
								S_BUF.BUFFER[x] := BYTE#16#31;
								x := x + 1;
								S_BUF.BUFFER[x] := BYTE#16#3B;
							END_IF;
							IF (FRONT_COLOR AND BYTE#2#00010000) > BYTE#0 THEN
								x := x + 1;
								S_BUF.BUFFER[x] := BYTE#16#35;
								x := x + 1;
								S_BUF.BUFFER[x] := BYTE#16#3B;
							END_IF;
						END_IF;
						x := x + 1;
						S_BUF.BUFFER[x] := BYTE#16#33;
						x := x + 1;
						S_BUF.BUFFER[x] := (FRONT_COLOR AND BYTE#2#00000111) OR BYTE#16#30;
						x := x + 1;
						S_BUF.BUFFER[x] := BYTE#16#6D;
						last_FC := FRONT_COLOR;
					END_IF;

					IF X_POS > BYTE#0 AND Y_POS > BYTE#0 THEN
						x := x + 1;
						S_BUF.BUFFER[x] := BYTE#16#1B;
						x := x + 1;
						S_BUF.BUFFER[x] := BYTE#16#5B;
						x := x + 1;
						S_BUF.BUFFER[x] := SHR(INT_TO_BCDC(BYTE_TO_INT(Y_POS)),4) OR BYTE#16#30;
						x := x + 1;
						S_BUF.BUFFER[x] := (INT_TO_BCDC(BYTE_TO_INT(Y_POS)) AND BYTE#16#0F) OR BYTE#16#30;
						x := x + 1;
						S_BUF.BUFFER[x] := BYTE#16#3B;
						x := x + 1;
						S_BUF.BUFFER[x] := SHR(INT_TO_BCDC(BYTE_TO_INT(X_POS)),4) OR BYTE#16#30;
						x := x + 1;
						S_BUF.BUFFER[x] := (INT_TO_BCDC(BYTE_TO_INT(X_POS)) AND BYTE#16#0F) OR BYTE#16#30;
						x := x + 1;
						S_BUF.BUFFER[x] := BYTE#16#48;
					END_IF;

					IF LEN(TEXT) > 0 THEN
						_STRING_TO_BUFFER(str:=TEXT,pos:=x + 1,size:=s_buf_size,pt:=S_BUF.BUFFER);
						S_BUF.BUFFER:=_STRING_TO_BUFFER.pt;
						x := x + LEN(TEXT);
					END_IF;

					IF b3_cr_lr THEN
						x := x + 1;
						S_BUF.BUFFER[x] := BYTE#16#0D;
						x := x + 1;
						S_BUF.BUFFER[x] := BYTE#16#0A;
					END_IF;

					DONE := TRUE;

					IF b7_no_flush THEN
						S_BUF.SIZE := INT_TO_UINT(x + 1);
						x := -1;
					END_IF;
				END_IF;
			END_IF;
		END_IF;
	END_CASE;

	IP_FIFO(FIFO:=IP_C.FIFO,STATE:=IP_STATE,ID:=IP_ID);
	IP_C.FIFO:=IP_FIFO.FIFO;
	IP_STATE := IP_FIFO.STATE;
	IP_ID:=IP_FIFO.ID;

	READY := IP_C.C_STATE > BYTE#127;
	DONE := FALSE;

	CASE state OF

	00:
		IF ENABLE THEN
			state := 10;
			IP_STATE := BYTE#1;
		END_IF;

	10:
		IF IP_STATE = BYTE#3 THEN

			IP_C.C_PORT     := WORD#23;
			IP_C.C_IP       := DWORD#00;
			IP_C.C_MODE     := BYTE#4;
			IP_C.TIME_RESET := TRUE;
			IP_C.C_ENABLE   := TRUE;
			IP_C.R_OBSERVE  := FALSE;
			state := 20;
		END_IF;

	20: IF IP_C.ERROR > DWORD#0 THEN
			IP_C.TIME_RESET := TRUE;
		END_IF;
		IF S_BUF.SIZE = UINT#0 THEN
			IF NOT ENABLE THEN
				IP_STATE := BYTE#4;
				IP_C.C_ENABLE := FALSE;
				state := 0;
			END_IF;
			IF IP_C.C_STATE = BYTE#1  THEN
				INIT := FALSE;
			ELSIF READY THEN
				IF IP_C.C_STATE = BYTE#254 AND NOT INIT THEN
					INIT := TRUE;
					last_FC := NOT FRONT_COLOR;

					_STRING_TO_BUFFER(str:='#[?7h#[0;3#;4#m#[2J',pos:=0,size:=S_BUF_SIZE,pt:=S_BUF.BUFFER);
					S_BUF.BUFFER:=_STRING_TO_BUFFER.pt;

					S_BUF.BUFFER[0] := BYTE#16#1B;
					IF (OPTION AND BYTE#2#0000_0010) > BYTE#0 THEN
						S_BUF.BUFFER[4] := BYTE#16#6C;
					END_IF;
					x := 4;
					IF (OPTION AND BYTE#2#0000_0001) > BYTE#0 THEN

						S_BUF.BUFFER[05] := BYTE#16#1B;
						S_BUF.BUFFER[10] := (FRONT_COLOR AND BYTE#2#00000111) OR BYTE#16#30;
						S_BUF.BUFFER[13] := (BACK_COLOR AND BYTE#2#00000111) OR BYTE#16#30;
						S_BUF.BUFFER[15] := BYTE#16#1B;
						x := 18;
					ELSE
						x := x + 1;
						S_BUF.BUFFER[x] := BYTE#16#0A;
					END_IF;
				END_IF;

				IF (INT_TO_UINT(x + LEN(TEXT) + 21) > S_BUF_SIZE) OR (x >= 0 AND NOT SEND) THEN
					S_BUF.SIZE := INT_TO_UINT(x + 1);
					x := -1;
				ELSIF SEND THEN

					IF (OPTION AND BYTE#2#0000_0100) > BYTE#0 AND FRONT_COLOR <> last_FC THEN
						x := x + 1;
						S_BUF.BUFFER[x] := BYTE#16#1B;
						x := x + 1;
						S_BUF.BUFFER[x] := BYTE#16#5B;
						IF ((FRONT_COLOR AND BYTE#2#0001_1000) XOR (last_FC AND BYTE#2#0001_1000)) <> BYTE#00 OR TRUE THEN
							x := x + 1;
							S_BUF.BUFFER[x] := BYTE#16#30;
							x := x + 1;
							S_BUF.BUFFER[x] := BYTE#16#3B;
							IF (FRONT_COLOR AND BYTE#2#00001000) = BYTE#0 THEN
								x := x + 1;
								S_BUF.BUFFER[x] := BYTE#16#31;
								x := x + 1;
								S_BUF.BUFFER[x] := BYTE#16#3B;
							END_IF;
							IF (FRONT_COLOR AND BYTE#2#00010000) > BYTE#0 THEN
								x := x + 1;
								S_BUF.BUFFER[x] := BYTE#16#35;
								x := x + 1;
								S_BUF.BUFFER[x] := BYTE#16#3B;
							END_IF;
						END_IF;
						x := x + 1;
						S_BUF.BUFFER[x] := BYTE#16#33;
						x := x + 1;
						S_BUF.BUFFER[x] := (FRONT_COLOR AND BYTE#2#00000111) OR BYTE#16#30;
						x := x + 1;
						S_BUF.BUFFER[x] := BYTE#16#6D;
						last_FC := FRONT_COLOR;
					END_IF;

					IF X_POS > BYTE#0 AND Y_POS > BYTE#0 THEN
						x := x + 1;
						S_BUF.BUFFER[x] := BYTE#16#1B;
						x := x + 1;
						S_BUF.BUFFER[x] := BYTE#16#5B;
						x := x + 1;
						S_BUF.BUFFER[x] := SHR_BYTE(INT_TO_BCDC(_BYTE_TO_INT(Y_POS)),4) OR BYTE#16#30;
						x := x + 1;
						S_BUF.BUFFER[x] := (INT_TO_BCDC(_BYTE_TO_INT(Y_POS)) AND BYTE#16#0F) OR BYTE#16#30;
						x := x + INT#1;
						S_BUF.BUFFER[x] := BYTE#16#3B;
						x := x + 1;
						S_BUF.BUFFER[x] := SHR_BYTE(INT_TO_BCDC(_BYTE_TO_INT(X_POS)),4) OR BYTE#16#30;
						x := x + 1;
						S_BUF.BUFFER[x] := (INT_TO_BCDC(_BYTE_TO_INT(X_POS)) AND BYTE#16#0F) OR BYTE#16#30;
						x := x + 1;
						S_BUF.BUFFER[x] := BYTE#16#48;
					END_IF;

					IF LEN(TEXT) > 0 THEN

						_STRING_TO_BUFFER(str:=TEXT,pos:=x + 1,size:=S_BUF_SIZE,pt:=S_BUF.BUFFER);
						S_BUF.BUFFER:=_STRING_TO_BUFFER.pt;
						x := x + LEN(TEXT);
					END_IF;

					IF (OPTION AND BYTE#2#0000_1000) > BYTE#0 THEN
						x := x + 1;
						S_BUF.BUFFER[x] := BYTE#16#0D;
						x := x + 1;
						S_BUF.BUFFER[x] := BYTE#16#0A;
					END_IF;

					DONE := TRUE;

					IF (OPTION AND BYTE#2#1000_0000) = BYTE#0 THEN
						S_BUF.SIZE := INT_TO_UINT(x + 1);
						x := -1;
					END_IF;
				END_IF;
			END_IF;
		END_IF;
	END_CASE;

	IP_FIFO(FIFO:=IP_C.FIFO,STATE:=IP_STATE,ID:=IP_ID);
	IP_C.FIFO:=IP_FIFO.FIFO;
	IP_STATE := IP_FIFO.STATE;
	IP_ID:=IP_FIFO.ID;

END_FUNCTION_BLOCK

PROGRAM program0
	VAR
		TEXT :	oscat_STRING250;
		ENABLE :	BOOL;
		SEND :	BOOL;
		OPTION :	BYTE;
		BACK_COLOR :	BYTE;
		FRONT_COLOR :	BYTE;
		X_POS :	BYTE;
		Y_POS :	BYTE;
		PORT :	WORD := WORD#23;
		IP_C :	oscat_IP_C;
		S_BUF :	oscat_NETWORK_BUFFER;
		READY :	BOOL;
		DONE :	BOOL;

		func_block : TELNET_PRINT_Block;
	END_VAR
	func_block.TEXT := TEXT;
	func_block.ENABLE := ENABLE;
	func_block.SEND := SEND;
	func_block.OPTION := OPTION;
	func_block.BACK_COLOR := BACK_COLOR;
	func_block.FRONT_COLOR := FRONT_COLOR;
	func_block.X_POS := X_POS;
	func_block.Y_POS := Y_POS;
	func_block.PORT := PORT;
	func_block.IP_C := IP_C;
	func_block.S_BUF := S_BUF;

	func_block();
	IP_C  := func_block.IP_C;
	S_BUF  := func_block.S_BUF;
	READY  := func_block.READY;
	DONE  := func_block.DONE;
END_PROGRAM

CONFIGURATION Config0
	RESOURCE Res0 ON PLC
		TASK task0(INTERVAL := T#20ms,PRIORITY := 0);
		PROGRAM instance0 WITH task0 : program0;
	END_RESOURCE
END_CONFIGURATION

(* ---- 741-MB_SERVER.ST ---- *)
TYPE
	oscat_IP_FIFO128_DATA  : ARRAY [1..128] OF BYTE;
	oscat_Mailbox  : ARRAY [1..16] OF BYTE;

	oscat_NW_BUF_SHORT : ARRAY [0..1407] OF BYTE;
	oscat_NW_BUF_LONG  : ARRAY [0..4095] OF BYTE;

	oscat_IP_FIFO_DATA :
	STRUCT
		X       : oscat_IP_FIFO128_DATA; (* IP_ID FIFO Speicher          *)
		Y       : oscat_IP_FIFO128_DATA; (* IP_ID Z�hler                 *)
		ID      : BYTE;                  (* h�chste vergabene id         *)
		MAX_ID  : BYTE;                  (* maximal Anmeldungen pro ID   *)
		INIT    : BOOL;                  (* Initialisierung durchgef�hrt *)
		EMPTY   : BOOL;                  (* FIFO leer                    *)
		FULL    : BOOL;                  (* FIFO voll                    *)
		TOP     : INT;                   (* maximale anzahl in FIFO      *)
		NW      : INT;                   (* Schreibzeiger                *)
		NR      : INT;                   (* Lesezeiger                   *)
	END_STRUCT;

	oscat_IP_C:
	STRUCT
		C_MODE:			BYTE;          		(*W Mode: TCP/UCP AKTIV/PASSIV                               *)
		C_PORT:         WORD;          		(*W Portnummer                                               *)
		C_IP:           DWORD;         		(*W IP-Adresse gepackt wwxxyyzz = www.xxx.yyy.zzz            *)
		C_STATE:        BYTE;          		(*R Verbindungsstatus ON/OFF + Flanke ON/OFF                 *)
		C_ENABLE:       BOOL;          		(*W Freigabe f�r Connect                                     *)
		R_OBSERVE:      BOOL;          		(*W Empfang ueberwachen                                      *)
		TIME_RESET:     BOOL;          		(*W Alle Timer ruecksetzen                                   *)
		ERROR:          DWORD;         		(*R vvwwxxyy (vv = CON_ERROR, ww = SEN_ERROR, xx = REC_ERROR *)
		FIFO:           oscat_IP_FIFO_DATA; (*I IP FIFO Struktur                                         *)
		MAILBOX:		oscat_Mailbox;		(*I Mailbox: Datenbereich f�r Bausteindatenaustausch         *)
	END_STRUCT;

	oscat_NETWORK_BUFFER :
	STRUCT
		SIZE   : UINT;
		BUFFER : oscat_NW_BUF_LONG;
	END_STRUCT;

	oscat_NETWORK_BUFFER_SHORT :
	STRUCT
	SIZE   : UINT;
	BUFFER : oscat_NW_BUF_SHORT;
	END_STRUCT;

	oscat_aW0_255	: ARRAY [0..255] OF WORD;
	oscat_VMAP_DATA :
	STRUCT
		FC       : DWORD;
		V_ADR    : INT;
		V_SIZE   : INT;
		P_ADR    : INT;
		TIME_OUT : TIME;
	END_STRUCT;

	oscat_MB_VMAP : ARRAY [1..10] OF oscat_VMAP_DATA;

	csv_parser_demo_col : ARRAY [1..4] OF REAL;
	csv_parser_demo     : ARRAY [1..2] OF csv_parser_demo_col;

END_TYPE

FUNCTION_BLOCK MB_VMAP_Block

	VAR_IN_OUT
		VMAP :	oscat_MB_VMAP;
	END_VAR

	VAR_INPUT
		FC :	INT;
		V_ADR :	INT;
		V_CNT :	INT;
		SIZE :	INT;
	END_VAR

	VAR_OUTPUT
		P_ADR :	INT;
		P_BIT :	INT;
		ERROR :	BYTE;
	END_VAR

	VAR
		i :	INT;
		vopt :	DWORD;
		vadr :	INT;
		padr :	INT;
		mask :	DWORD;
		vsize :	INT;
		w_tmp :	WORD;
		i_tmp :	INT;
		init :	BOOL;
	END_VAR

	IF init = FALSE THEN
		init := TRUE;
		IF VMAP[1].FC = DWORD#0 THEN
			VMAP[1].FC := DWORD#16#FFFF_FFFF;
			VMAP[1].V_ADR := 0;
			VMAP[1].V_SIZE := 256;
			VMAP[1].P_ADR := 0;
		END_IF;
	END_IF;

	ERROR := BYTE#02;
	mask := SHL(DWORD#1,FC);

	IF (mask AND DWORD#2#00000000_01000000_00000000_01100000) <> DWORD#0 THEN
		V_CNT := 1;
	ELSIF V_CNT = 0 THEN
		RETURN;
	END_IF;

	FOR i := 1 TO 10 DO
		vopt := VMAP[i].FC;
		IF (vopt AND mask) <> DWORD#0 THEN
			vadr := VMAP[i].V_ADR;
			vsize := VMAP[i].V_SIZE;
			padr := VMAP[i].P_ADR;

			IF (mask AND DWORD#2#00000000_00000000_10000000_00100110) <> DWORD#0 THEN
				i_tmp := WORD_TO_INT(SHR(INT_TO_WORD(V_ADR + V_CNT -1),4))+1;
				IF i_tmp <= SIZE AND i_tmp <= vsize THEN
					w_tmp := INT_TO_WORD(V_ADR);
					P_ADR := WORD_TO_INT(SHR(w_tmp,4)) + padr;
					P_BIT := WORD_TO_INT(w_tmp AND WORD#16#000F);
					ERROR := BYTE#0;
					EXIT;
				END_IF;
			ELSIF (mask AND DWORD#2#00000000_11000001_00000000_01011000) <> DWORD#0 THEN
				IF V_ADR >= vadr AND V_ADR + V_CNT <= vadr + vsize THEN
					P_ADR := V_ADR - vadr + padr;
					IF P_ADR + V_CNT <= SIZE THEN
						ERROR := BYTE#0;
						EXIT;
					END_IF;
				END_IF;
			ELSE
				ERROR := BYTE#01;
				RETURN;
			END_IF;
		END_IF;
	END_FOR;

	IF ERROR = BYTE#0 THEN
		IF (mask AND DWORD#2#00000000_11000001_10000000_01100000) <> DWORD#0 THEN
			VMAP[i].TIME_OUT := T#1ms;
		END_IF;
	END_IF;

END_FUNCTION_BLOCK

FUNCTION _BYTE_TO_INT:INT
	VAR_INPUT
		IN :	BYTE;
	END_VAR

	_BYTE_TO_INT := USINT_TO_INT(BYTE_TO_USINT(IN));
END_FUNCTION

FUNCTION_BLOCK IP_FIFO_Block

  VAR_IN_OUT
    FIFO :	oscat_IP_FIFO_DATA;
    ID :	BYTE;
    STATE :	BYTE;
  END_VAR

  VAR
    tmp :	INT;
  END_VAR

  IF NOT FIFO.INIT THEN
    FIFO.INIT		:= TRUE;
    FIFO.NW		:= 1;
    FIFO.NR		:= 1;
    FIFO.EMPTY	:= TRUE;
    FIFO.FULL		:= FALSE;
    FIFO.TOP		:= 128;
    FIFO.MAX_ID	:= BYTE#1;
  END_IF;

  IF ID = BYTE#00 THEN
    IF FIFO.ID < INT_TO_BYTE(FIFO.TOP) THEN
      ID := USINT_TO_BYTE(BYTE_TO_USINT(FIFO.ID) + USINT#1);
      FIFO.ID := ID ;

    ELSIF STATE < BYTE#200 THEN
      STATE := BYTE#255;
    RETURN;
    END_IF;
  END_IF;

  IF STATE = BYTE#1 AND NOT FIFO.FULL THEN
    tmp := _BYTE_TO_INT(ID);
    IF FIFO.Y[tmp] < FIFO.MAX_ID THEN
      FIFO.Y[tmp] := USINT_TO_BYTE(BYTE_TO_USINT(FIFO.Y[tmp]) + USINT#1);
      tmp := FIFO.NW;
      FIFO.X[tmp] := ID;
      IF FIFO.NW = FIFO.TOP THEN FIFO.NW := 1; ELSE FIFO.NW := FIFO.NW + 1; END_IF;
      FIFO.FULL := FIFO.NW = FIFO.NR;
    FIFO.EMPTY := FALSE;
      STATE := BYTE#2;
    END_IF;
  END_IF;

  IF STATE = BYTE#2 AND NOT FIFO.EMPTY THEN
    tmp := FIFO.NR;
    IF ID = FIFO.X[tmp] THEN
      STATE := BYTE#3;
    END_IF;
  END_IF;

  IF STATE = BYTE#4 AND NOT FIFO.EMPTY THEN

    tmp := FIFO.NR;
    IF ID = FIFO.X[tmp] THEN
      tmp := _BYTE_TO_INT(ID);
      FIFO.Y[tmp] := USINT_TO_BYTE(BYTE_TO_USINT(FIFO.Y[tmp]) - USINT#1);

      IF FIFO.NR = FIFO.TOP THEN FIFO.NR := 1; ELSE FIFO.NR := FIFO.NR + 1; END_IF;
      FIFO.EMPTY := FIFO.NR = FIFO.NW;
    FIFO.FULL := FALSE;
    END_IF;
    STATE := BYTE#5;
  END_IF;

END_FUNCTION_BLOCK

FUNCTION _UDINT_TO_TIME:TIME

	VAR_INPUT
		IN :	UDINT;
	END_VAR

	_UDINT_TO_TIME := DINT_TO_TIME(UDINT_TO_DINT(IN));

END_FUNCTION

FUNCTION_BLOCK T_PLC_MS_block

	VAR_OUTPUT
		T_PLC_MS :	UDINT;
	END_VAR

	VAR_EXTERNAL
		PLC_TICKS_PER_SEC :	INT;
		PLC_SYS_TICK_CNT :	DINT;
	END_VAR

	VAR
		debug :	BOOL;(*Debug-Mode ON / OFF*)
		N :	INT;(*Debug-Faktor*)
		Offset :	UDINT;(*Debug-Offset*)
		temp :	DWORD := DWORD#1;(*Debug-Offset*)
		mode :	BOOL;(*modus*)
		faktor :	UDINT;(*Systemtakt-Faktor*)
		init :	BOOL;
		v_plc_ticks_per_sec :	UDINT;
		base :	UDINT := UDINT#1000;
	END_VAR

	IF init = FALSE THEN
		v_plc_ticks_per_sec := INT_TO_UDINT(PLC_TICKS_PER_SEC);
		IF v_plc_ticks_per_sec = UDINT#1024 THEN
			faktor := UDINT#1;
			mode := FALSE;
		ELSIF v_plc_ticks_per_sec > UDINT#0 THEN
			IF v_plc_ticks_per_sec <= base THEN
				faktor := base / v_plc_ticks_per_sec;
				mode := FALSE;
			ELSE
				faktor := v_plc_ticks_per_sec / base;
				mode := TRUE;
			END_IF;
		ELSE
			faktor := UDINT#1;
		END_IF;
		init := TRUE;
	END_IF;

	IF mode THEN
		T_PLC_MS := DINT_TO_UDINT(PLC_SYS_TICK_CNT) / faktor;
	ELSE
		T_PLC_MS := DINT_TO_UDINT(PLC_SYS_TICK_CNT) * faktor;
	END_IF;

	IF debug THEN
		T_PLC_MS := (DWORD_TO_UDINT(SHL(UDINT_TO_DWORD(T_PLC_MS),N) OR SHL(temp,N)) - UDINT#1) + Offset;
	END_IF;

END_FUNCTION_BLOCK

FUNCTION WORD_OF_BYTE:WORD
	VAR_INPUT
		B1 :	BYTE;
		B0 :	BYTE;
	END_VAR
	WORD_OF_BYTE := SHL(BYTE_TO_WORD(B1),8) OR BYTE_TO_WORD(B0);
END_FUNCTION

FUNCTION BIT_LOAD_W:WORD
	VAR_INPUT
		IN :	WORD;
		VAL :	BOOL;
		POS :	INT;
	END_VAR

	IF VAL THEN
		BIT_LOAD_W := in OR SHL(WORD#1,pos);
	ELSE
		BIT_LOAD_W := in AND (NOT SHL(WORD#1,pos));
	END_IF;
END_FUNCTION

FUNCTION_BLOCK MB_SERVER_Block

	VAR_IN_OUT
		IP_C :	oscat_IP_C;
		S_BUF :	oscat_NETWORK_BUFFER_SHORT;
		R_BUF :	oscat_NETWORK_BUFFER_SHORT;
		VMAP :	oscat_MB_VMAP;
		DATA :	oscat_aW0_255;
	END_VAR

	VAR_INPUT
		DATA_SIZE :	INT;
		ENABLE :	BOOL;
		UDP :	BOOL;
	END_VAR

	VAR_OUTPUT
		ERROR :	DWORD;
	END_VAR

	VAR
		MB_VMAP :	MB_VMAP_Block;
		adr1 :	INT;
		adr2 :	INT;
		points :	INT;
		points2 :	INT;
		coils :	BYTE;
		mask :	BYTE;
		idx1 :	INT;
		idx2 :	INT;
		bit_pos :	INT;
		count :	INT;
		fc :	INT;
		i :	INT;
		state :	INT;
		IP_STATE :	BYTE;
		IP_ID :	BYTE;
		IP_FIFO :	IP_FIFO_Block;
		w_tmp :	WORD;
		last_cycle :	TIME;
		tx :	TIME;
		T_PLC_MS :	T_PLC_MS_Block;
		t :	TON;
		ip_error :	BOOL;
	END_VAR

	T_PLC_MS();
	tx := UDINT_TO_TIME(T_PLC_MS.T_PLC_MS);

	FOR i := 1 TO 10 DO
		IF VMAP[i].TIME_OUT > T#0s THEN
			VMAP[i].TIME_OUT := VMAP[i].TIME_OUT + tx - last_cycle;
		END_IF;
	END_FOR;
	last_cycle := tx;
	ip_error := IP_C.ERROR > DWORD#0;

	CASE state OF

	00:
		IF ENABLE THEN
			state := 10;
			IP_STATE := BYTE#1;
		END_IF;

	10:
		IF IP_STATE = BYTE#3 THEN

			IP_C.C_PORT     := WORD#0;
			IP_C.C_IP       := DWORD#0;
			IP_C.C_MODE     := SEL(UDP,BYTE#4,BYTE#5);
			IP_C.TIME_RESET := TRUE;
			IP_C.C_ENABLE   := TRUE;
			IP_C.R_OBSERVE  := FALSE;
			state := 20;
		END_IF;

	20:	IF NOT ip_error THEN
			IF S_BUF.SIZE = UINT#0 AND R_BUF.SIZE > UINT#6 THEN
				IF  R_BUF.SIZE = WORD_TO_UINT(WORD_OF_BYTE(R_BUF.BUFFER[4],R_BUF.BUFFER[5])) + UINT#6 THEN
					ERROR := DWORD#00;

					FOR i := 0 TO 13 DO
						S_BUF.BUFFER[i] := R_BUF.BUFFER[i];
					END_FOR;

					fc := _BYTE_TO_INT(R_BUF.BUFFER[7]);

					adr1 := WORD_TO_INT(WORD_OF_BYTE(R_BUF.BUFFER[8],R_BUF.BUFFER[9]));
					points := WORD_TO_INT(WORD_OF_BYTE(R_BUF.BUFFER[10],R_BUF.BUFFER[11]));

					MB_VMAP(VMAP:=VMAP,FC:=fc,V_ADR:=adr1,V_CNT:=points,SIZE:=DATA_SIZE);
					VMAP:=MB_VMAP.VMAP;
					adr1:=MB_VMAP.P_ADR;
					bit_pos:=MB_VMAP.P_BIT;
					ERROR:=BYTE_TO_DWORD(MB_VMAP.ERROR);

					IF ERROR = DWORD#0 THEN
						CASE fc OF

						1..2 :
							count := 9;
							coils := BYTE#0;
							mask := BYTE#1;
							FOR i := 1 TO points DO
								IF mask = BYTE#0 THEN
									mask := BYTE#1;
									S_BUF.BUFFER[count] := coils;
									coils := BYTE#0;
									count := count + 1;
								END_IF;
								IF (DATA[adr1] AND SHL(WORD#1,bit_pos)) > WORD#0 THEN
									coils := coils OR mask;
								END_IF;

								bit_Pos := bit_Pos + 1;
								IF bit_pos > 15 THEN
									adr1 := adr1 + 1;
									bit_pos := 0;
								END_IF;

								mask := SHL(mask,1);
							END_FOR;
							S_BUF.BUFFER[Count] := coils;

							S_BUF.BUFFER[8] := INT_TO_BYTE(count - 8);
							S_BUF.SIZE := INT_TO_UINT(count + 1);

						3..4 :
							idx1 := 07;
							count := adr1 + points - 1;
							FOR i := adr1 TO count DO
								idx1 := idx1 + 2;
								idx2 := idx1 + 1;
								w_tmp := DATA[i];
								S_BUF.BUFFER[idx1] := WORD_TO_BYTE(SHR(w_tmp,8));
								S_BUF.BUFFER[idx2] := WORD_TO_BYTE(w_tmp);
							END_FOR;
							S_BUF.BUFFER[8] := SHL(INT_TO_BYTE(points),1);
							S_BUF.SIZE := INT_TO_UINT(idx2 + 1);
						5 :
							DATA[adr1]:=BIT_LOAD_W(DATA[adr1],R_BUF.BUFFER[10]>BYTE#0,bit_pos);
							S_BUF.SIZE := UINT#12;
						6 :
							DATA[adr1] := WORD_OF_BYTE(R_BUF.BUFFER[10],R_BUF.BUFFER[11]);
							S_BUF.SIZE := UINT#12;
						15 :
							mask := BYTE#1;
							idx1 := 13;
							FOR i := 1 TO points DO
								DATA[adr1]:=BIT_LOAD_W(DATA[adr1],(R_BUF.BUFFER[idx1] AND mask)>BYTE#0,bit_pos);
								bit_pos := bit_pos + 1;
								IF bit_pos > 15 THEN
									adr1 := adr1 + 1;
									bit_pos := 0;
								END_IF;
								mask := ROL(mask,1);
								IF mask = BYTE#1 THEN
									idx1 := idx1 +1;
								END_IF;
							END_FOR;
							S_BUF.SIZE := UINT#12;
						16 :
							idx1 := 11;
							count := adr1 + points -1;
							FOR i := adr1 TO Count DO
								idx1 := idx1 + 2;
								idx2 := idx1 + 1;
								Data[i] := WORD_OF_BYTE(R_BUF.BUFFER[idx1],R_BUF.BUFFER[idx2]);
							END_FOR;
							S_BUF.SIZE := UINT#12;
						22 :
							w_tmp := WORD_OF_BYTE(R_BUF.BUFFER[11],R_BUF.BUFFER[11]);
							DATA[adr1] := (DATA[adr1] AND w_tmp) OR (WORD_OF_BYTE(R_BUF.BUFFER[12],R_BUF.BUFFER[13]) AND (NOT w_tmp));
							S_BUF.SIZE := UINT#14;
						23 :
							adr2 := WORD_TO_INT(WORD_OF_BYTE(R_BUF.BUFFER[12],R_BUF.BUFFER[13]));
							points2 := WORD_TO_INT(WORD_OF_BYTE(R_BUF.BUFFER[14],R_BUF.BUFFER[15]));

							MB_VMAP(VMAP:=VMAP,FC:=16,V_ADR:=adr2,V_CNT:=points2,SIZE:=DATA_SIZE);
							VMAP:=MB_VMAP.VMAP;
							adr2:=MB_VMAP.P_ADR;
							ERROR:=BYTE_TO_DWORD(MB_VMAP.ERROR);

							IF ERROR = DWORD#0 THEN
								idx1 := 15;
								count := adr2 + points2 -1;
								FOR i := adr2 TO count DO
									idx1 := idx1 + 2;
									idx2 := idx1 + 1;
									Data[i] := WORD_OF_BYTE(R_BUF.BUFFER[idx1],R_BUF.BUFFER[idx2]);
								END_FOR;

								idx1 := 07;
								count := adr1 + points - 1;
								FOR i := adr1 TO count DO
									idx1 := idx1 + 2;
									idx2 := idx1 + 1;
									w_tmp := DATA[i];
									S_BUF.BUFFER[idx1] := WORD_TO_BYTE(SHR(w_tmp,8));
									S_BUF.BUFFER[idx2] := WORD_TO_BYTE(w_tmp);
								END_FOR;
								S_BUF.BUFFER[8] := SHL(INT_TO_BYTE(points),1);
								S_BUF.SIZE := INT_TO_UINT(idx2 + 1);

							END_IF;

						ELSE
							ERROR := DWORD#01;
						END_CASE;
					END_IF;
				END_IF;

				IF ERROR > DWORD#0 THEN
					S_BUF.BUFFER[7] := S_BUF.BUFFER[7] OR BYTE#2#1000_0000;
					S_BUF.BUFFER[8] := DWORD_TO_BYTE(ERROR);
					S_BUF.SIZE := UINT#9;
				END_IF;

				S_BUF.BUFFER[4] := BYTE#0;
				S_BUF.BUFFER[5] := UINT_TO_BYTE(S_BUF.SIZE - UINT#6);

			END_IF;
		ELSE
			ERROR := IP_C.ERROR;
		END_IF;

		t(IN:= ip_error, PT:=T#5s);
		IF t.Q THEN
			IP_C.TIME_RESET := TRUE;
		END_IF;

		R_BUF.SIZE := UINT#0;

		IF ENABLE = FALSE THEN
			IP_STATE := BYTE#4;
			state := 00;
		END_IF;
	END_CASE;

	IP_FIFO(FIFO:=IP_C.FIFO,STATE:=IP_STATE,ID:=IP_ID);
	IP_C.FIFO:=IP_FIFO.FIFO;
	IP_STATE := IP_FIFO.STATE;
	IP_ID:=IP_FIFO.ID;

END_FUNCTION_BLOCK

PROGRAM program0
	VAR
		IP_C :	oscat_IP_C;
		S_BUF :	oscat_NETWORK_BUFFER_SHORT;
		R_BUF :	oscat_NETWORK_BUFFER_SHORT;
		VMAP :	oscat_MB_VMAP;
		DATA :	oscat_aW0_255;
		DATA_SIZE :	INT;
		ENABLE :	BOOL;
		UDP :	BOOL;
		ERROR :	DWORD;

		func_block : MB_SERVER_Block;
	END_VAR
	func_block.IP_C := IP_C;
	func_block.S_BUF := S_BUF;
	func_block.R_BUF := R_BUF;
	func_block.VMAP := VMAP;
	func_block.DATA := DATA;
	func_block.DATA_SIZE := DATA_SIZE;
	func_block.ENABLE := ENABLE;
	func_block.UDP := UDP;

	func_block();
  	IP_C  := func_block.IP_C;
	S_BUF  := func_block.S_BUF;
	R_BUF  := func_block.R_BUF;
	VMAP  := func_block.VMAP;
	DATA  := func_block.DATA;
	ERROR  := func_block.ERROR;

END_PROGRAM

CONFIGURATION Config0

	VAR_GLOBAL
		PLC_TICKS_PER_SEC :	INT;
		PLC_SYS_TICK_CNT :	DINT;
	END_VAR

  	RESOURCE Res0 ON PLC
    	TASK task0(INTERVAL := T#20ms,PRIORITY := 0);
    	PROGRAM instance0 WITH task0 : program0;
  	END_RESOURCE

END_CONFIGURATION

(* ---- 10-ISC_NUM.ST ---- *)
FUNCTION ISC_NUM:BOOL

	VAR_INPUT
		IN :	BYTE;
	END_VAR

	ISC_NUM := IN > BYTE#47 AND IN < BYTE#58;

END_FUNCTION

PROGRAM program0
	VAR
		IN : BYTE;
		OUT : BOOL;
	END_VAR

	OUT := ISC_NUM(IN);
END_PROGRAM

CONFIGURATION Config0

	RESOURCE Res0 ON PLC
		TASK task0(INTERVAL := T#20ms,PRIORITY := 0);
		PROGRAM instance0 WITH task0 : program0;
	END_RESOURCE

END_CONFIGURATION
